// TIA Portal V17 export
// export: Created 2025-07-01T12:14:22.0161746Z, ExportSetting WithDefaults, DisplayName Totally Integrated Automation Portal, DisplayVersion V17, DisplayName TIA Portal Openness, DisplayVersion V17, DisplayName TIA Portal Version Control Interface, DisplayVersion V17, DisplayName SINAMICS Startdrive Advanced, DisplayVersion V17, DisplayName SINAMICS Startdrive G130, G150, S120, S150, SINAMICS MV, S210, DisplayVersion V17, DisplayName SINAMICS Startdrive G110M, G120, G120C, G120D, G120P, G115D, DisplayVersion V17, DisplayName STEP 7 Professional, DisplayVersion V17, DisplayName STEP 7 Safety, DisplayVersion V17, DisplayName WinCC Professional, DisplayVersion V17
FUNCTION_BLOCK "3PosLifter__Updated_V2_a4fa82_3a45ac7d-3c57-493c-83a9-58625a874be0 (2) - Copy_22ffb1"   // FB3, LAD
VERSION : 0.1
// stored: AutoNumber true, IsIECCheckEnabled false, UDAEnableTagReadback false
   VAR_INPUT
      iAreaClearConv : Bool;
      iAreaClearTransL2 : Bool;
      iAreaClear_TT : Bool;
      iAutoRunning : Bool;
      iErrorAck : Bool;
      iL1PalletPrsnt : Bool;
      iL1S1Raise : Bool;
      iL1S2Down : Bool;
      iL1S2DownOver : Bool;
      iL2PalletPrsent : Bool;
      iL2S1Down : Bool;
      iL2S1Raise : Bool;
      iL2s2DownOver : Bool;
      iL2s2Raise : Bool;
      iLiffterAtPos1 : Bool;
      iLiffterAtPos2 : Bool;
      iLiffterAtPos3 : Bool;
      iLiffterAtPos4 : Bool;
      iLifterAt1 : Bool;
      iLifterAtPos1 : Bool;
      iLifterAtPos2 : Bool;
      iLifterAtPos3 : Bool;
      iLifterAtPos4 : Bool;
      iOTSFrmConv : Bool;
      iPalAtTT : Bool;
      iPalletAtL1 : Bool;
      iPalletAtL2 : Bool;
      iPalletAtTT : Bool;
      iPalletPrsntL1 : Bool;
      iRTRFrmConv : Bool;
      iRTRFrmTT : Bool;
      iRTRFrm_TT : Bool;
      iReacvAreaClr : Bool;
      iReceiveAreaClear : Bool;
      iReceiveAreaClrConv : Bool;
      iRecvAreaClear : Bool;
      iReset_fault : Bool;
      iRunOutActive : Bool;
      iRunOutCycle : Bool;
      iSstMode : Bool;
      iSstPB : Bool;
      iTransAreaClearConv : Bool;
      iTransAreaClr : Bool;
      ipalletPrsntAtTT : Bool;
   END_VAR
   VAR_OUTPUT
      qL1S1Down : Bool;
      qL1S1raise : Bool;
      qL1S2Down : Bool;
      qL1S2Raise : Bool;
      qL1TrnsfrConv : Bool;
      qL2S1raise : Bool;
      qL2S2Down : Bool;
      qL2S2Raise : Bool;
      qLiffterAtPos2 : Bool;
      qLifterAtPos1 : Bool;
      qLifterAtPos3 : Bool;
      qLifterAtPos4 : Bool;
      qLifterGotoPos1 : Bool;
      qOTSToNext : Bool;
      qOTSTo_TT : Bool;
      qOutput1 : Bool;
      qRTRToConv : Bool;
      qRTRToTT : Bool;
      qRTR_To_Conv : Bool;
   END_VAR
   VAR_IN_OUT
      IqRx_Frm_TT : Bool;
      iqRx_frm_Conv : Bool;
      iqTX_To_Conv : Bool;
      iqTX_To_TT : Bool;
      iqTx_To_ConvPos4 : Bool;
      iqTx_To_Rej : Bool;
   END_VAR
   VAR DB_SPECIFIC
      StateNo : Int;
      s190_sStWtL1RcvComplete_T1 : Bool;
      s200_sStWtForL1StprUp_T1 : Bool;
      s240_sStWtL2TransComplete_T1 : Bool;
      s250_sStWtDeforkDone : Bool;
      s250_sStWtDeforkDone_Cond1 : Bool;
      s250_sStWtDeforkDone_Cond2 : Bool;
      s250_sStWtDeforkDone_T1 : Bool;
      sInitialConvRun : Bool;
      sInitialConvRun_T1 : Bool;
      sOTSTimeout : Bool;
      sSeq1Over : Bool;
      sSeq2Over : Bool;
      sSst : Bool;
      sSstPulse : Bool;
      sSstRise : Bool;
      sStChkPalAtTT : Bool;
      sStChkPalAtTT_T1 : Bool;
      sStChkPalAtTT_T2 : Bool;
      sStChkPalAtTT_T3 : Bool;
      sStChkPalletAtTT : Bool;
      sStChkPalletAtTT1 : Bool;
      sStChkPalletAtTT1_T1 : Bool;
      sStChkPalletAtTT1_T2 : Bool;
      sStChkPalletAtTT_T1 : Bool;
      sStChkPalletAtTT_T2 : Bool;
      sStChkPalletPrsntL1L2 : Bool;
      sStChkPalletPrsntL1L2_T1 : Bool;
      sStChkPalletPrsntL1L2_T2 : Bool;
      sStChkPalletPrsntL1L2_T3 : Bool;
      sStChkPalletPrsntL1L2_T4 : Bool;
      sStChkRunOutActive1 : Bool;
      sStChkRunOutActive1_T1 : Bool;
      sStChkRunOutActive1_T2 : Bool;
      sStL1S2Down : Bool;
      sStL1S2DownOver : Bool;
      sStL1S2DownOver_T1 : Bool;
      sStL1S2Down_T1 : Bool;
      sStNextRdyInTransit : Bool;
      sStNextRdyInTransit_1 : Bool;
      sStNextRdyInTransit_1_T1 : Bool;
      sStNextRdyInTransit_1_T2 : Bool;
      sStNextRdyInTransit_3 : Bool;
      sStNextRdyInTransit_3_T1 : Bool;
      sStNextRdyInTransit_3_T2 : Bool;
      sStNextRdyInTransit_T1 : Bool;
      sStNextRdyInTransit_T2 : Bool;
      sStRecovery : Bool;
      sStRecovery_T1 : Bool;
      sStRecovery_T2 : Bool;
      sStRecovery_T3 : Bool;
      sStRecovery_T4 : Bool;
      sStRecovery_T5 : Bool;
      sStRecovery_T6 : Bool;
      sStRecovery_T7 : Bool;
      sStRecovery_T8 : Bool;
      sStRunOutActive : Bool;
      sStRunOutActive_T1 : Bool;
      sStRunOutActive_T2 : Bool;
      sStWtDeforkDone : Bool;
      sStWtDeforkDone_T1 : Bool;
      sStWtForFaultReset : Bool;
      sStWtForFaultReset_T1 : Bool;
      sStWtForL1L2StoprsUp : Bool;
      sStWtForL1L2StoprsUp_T1 : Bool;
      sStWtForL1StprUp : Bool;
      sStWtForL1StprUp_T1 : Bool;
      sStWtL1PalRcvDone : Bool;
      sStWtL1PalRcvDone_T1 : Bool;
      sStWtL1RcvComplete : Bool;
      sStWtL1RcvComplete_T1 : Bool;
      sStWtL1RecvBegin : Bool;
      sStWtL1RecvBegin_T1 : Bool;
      sStWtL1S1Down1 : Bool;
      sStWtL1S1Down1_T1 : Bool;
      sStWtL1S2DownOver : Bool;
      sStWtL1S2DownOver_T1 : Bool;
      sStWtL1TransBegin : Bool;
      sStWtL1TransBeginPos4 : Bool;
      sStWtL1TransBeginPos4_T1 : Bool;
      sStWtL1TransBegin_T1 : Bool;
      sStWtL1TransComplet : Bool;
      sStWtL1TransComplet_T1 : Bool;
      sStWtL2RcvDone : Bool;
      sStWtL2RcvDone_T1 : Bool;
      sStWtL2RecvingActive : Bool;
      sStWtL2RecvingActive_T1 : Bool;
      sStWtL2S1Down : Bool;
      sStWtL2S1Down_T1 : Bool;
      sStWtL2S2Down : Bool;
      sStWtL2S2Down_T1 : Bool;
      sStWtL2TranBegin : Bool;
      sStWtL2TranBegin_T1 : Bool;
      sStWtL2TransComplete : Bool;
      sStWtL2TransComplete_T1 : Bool;
      sStWtLifterAtPos1 : Bool;
      sStWtLifterAtPos1_T1 : Bool;
      sStWtLifterAtPos2 : Bool;
      sStWtLifterAtPos2_T1 : Bool;
      sStWtLifterAtPos3 : Bool;
      sStWtLifterAtPos3_T1 : Bool;
      sStWtLifterAtPos4 : Bool;
      sStWtLifterAtPos4_T1 : Bool;
      sStWtLifterAtPosn1 : Bool;
      sStWtLifterAtPosn1_T1 : Bool;
      sStWtOTSFrmConv : Bool;
      sStWtOTSFrmConv1 : Bool;
      sStWtOTSFrmConv1_T1 : Bool;
      sStWtOTSFrmConv1_T2 : Bool;
      sStWtOTSFrmConv_T1 : Bool;
      sStWtOTSFrmTT : Bool;
      sStWtOTSFrmTT_T1 : Bool;
      sStWtRTRFrmConvPos4 : Bool;
      sStWtRTRFrmConvPos4_T1 : Bool;
      sStWtRTRFrmTT : Bool;
      sStWtRTRFrmTT_T1 : Bool;
      sStWtRcvBegin : Bool;
      sStWtRcvBegin_T1 : Bool;
      sStWtResetRel : Bool;
      sStWtResetRel_T1 : Bool;
      sStWtTransDonePos4 : Bool;
      sStWtTransDonePos4_T1 : Bool;
   END_VAR
   VAR_TEMP
      tOne : Bool;
   END_VAR
   VAR_TEMP   // added for the SCL form of the ladder/FBD networks
      _w1 : Bool;
   END_VAR
BEGIN

REGION Network 1
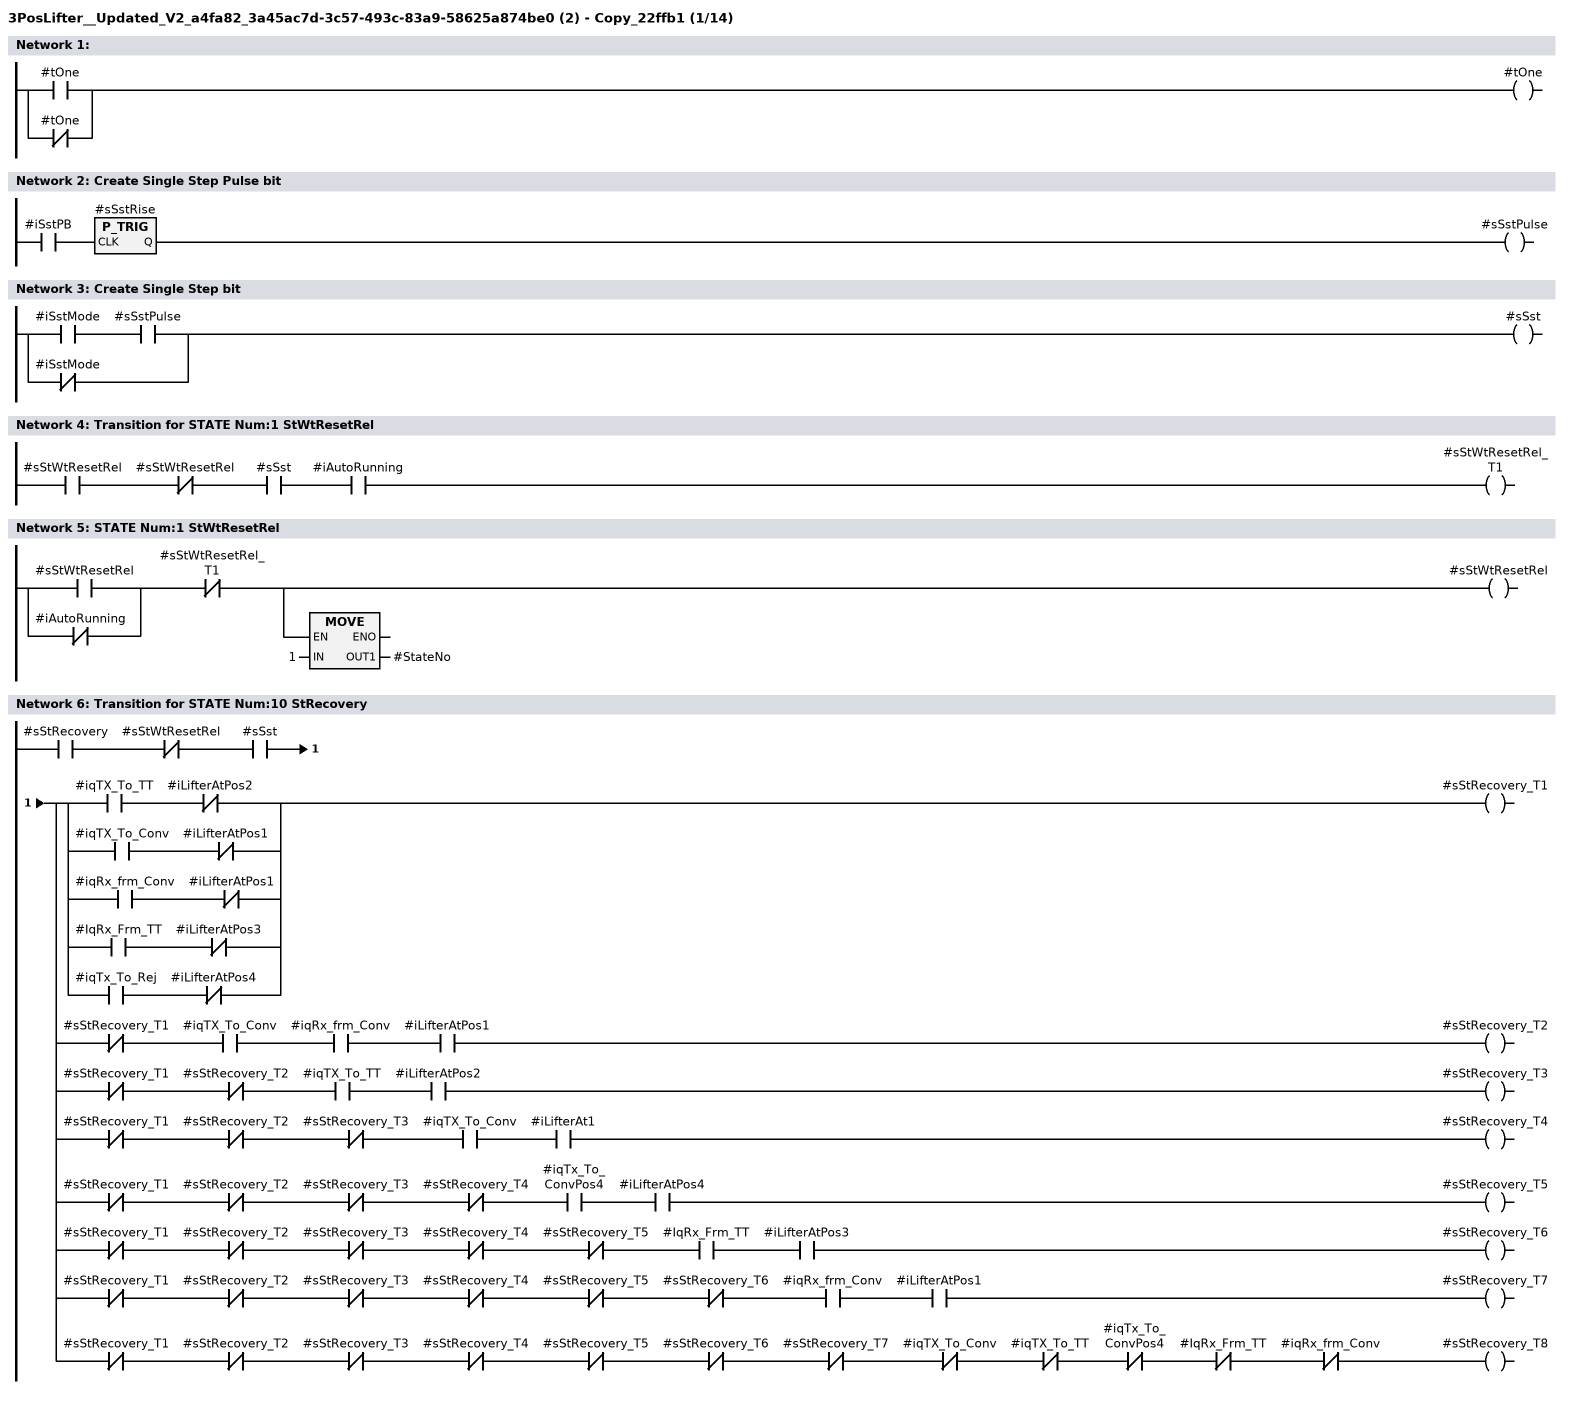
   RUNG wire#powerrail
      Contact( #tOne )
      wire#w1
      Coil( #tOne )
   END_RUNG
   RUNG wire#powerrail
      I_Contact( #tOne )
   END_RUNG wire#w1
   // the same network as SCL:
   #tOne := #tOne OR NOT #tOne;
END_REGION

REGION Network 2: Create Single Step Pulse bit
   RUNG wire#powerrail
      Contact( #iSstPB )
      P_Trig( #sSstRise )
      Coil( #sSstPulse )
   END_RUNG
   // the same network as SCL:
   #_w1 := #iSstPB AND NOT #sSstRise;   // rising edge
   #sSstRise := #iSstPB;
   #sSstPulse := #_w1;
END_REGION

REGION Network 3: Create Single Step bit
   RUNG wire#powerrail
      Contact( #iSstMode )
      Contact( #sSstPulse )
      wire#w1
      Coil( #sSst )
   END_RUNG
   RUNG wire#powerrail
      I_Contact( #iSstMode )
   END_RUNG wire#w1
   // the same network as SCL:
   #sSst := (#iSstMode AND #sSstPulse) OR NOT #iSstMode;
END_REGION

REGION Network 4: Transition for STATE Num:1 StWtResetRel
   RUNG wire#powerrail
      Contact( #sStWtResetRel )
      I_Contact( #sStWtResetRel )
      Contact( #sSst )
      Contact( #iAutoRunning )
      Coil( #sStWtResetRel_T1 )
   END_RUNG
   // the same network as SCL:
   #sStWtResetRel_T1 := #sStWtResetRel AND NOT #sStWtResetRel AND #sSst AND #iAutoRunning;
END_REGION

REGION Network 5: STATE Num:1 StWtResetRel
   RUNG wire#powerrail
      Contact( #sStWtResetRel )
      wire#w1
      I_Contact( #sStWtResetRel_T1 )
      wire#w2
      Coil( #sStWtResetRel )
   END_RUNG
   RUNG wire#powerrail
      I_Contact( #iAutoRunning )
   END_RUNG wire#w1
   RUNG wire#w2
      { S7_GenerateENO := "TRUE" } Move(in := 1, out1 => #StateNo)
   END_RUNG
   // the same network as SCL:
   #sStWtResetRel := (#sStWtResetRel OR NOT #iAutoRunning) AND NOT #sStWtResetRel_T1;
   IF #sStWtResetRel THEN #StateNo := 1; END_IF;
END_REGION

REGION Network 6: Transition for STATE Num:10 StRecovery
   RUNG wire#powerrail
      Contact( #sStRecovery )
      I_Contact( #sStWtResetRel )
      Contact( #sSst )
      wire#w1
      Contact( #iqTX_To_TT )
      I_Contact( #iLifterAtPos2 )
      wire#w2
      Coil( #sStRecovery_T1 )
   END_RUNG
   RUNG wire#w1
      Contact( #iqTX_To_Conv )
      I_Contact( #iLifterAtPos1 )
   END_RUNG wire#w2
   RUNG wire#w1
      Contact( #iqRx_frm_Conv )
      I_Contact( #iLifterAtPos1 )
   END_RUNG wire#w2
   RUNG wire#w1
      Contact( #IqRx_Frm_TT )
      I_Contact( #iLifterAtPos3 )
   END_RUNG wire#w2
   RUNG wire#w1
      Contact( #iqTx_To_Rej )
      I_Contact( #iLifterAtPos4 )
   END_RUNG wire#w2
   RUNG wire#w1
      I_Contact( #sStRecovery_T1 )
      Contact( #iqTX_To_Conv )
      Contact( #iqRx_frm_Conv )
      Contact( #iLifterAtPos1 )
      Coil( #sStRecovery_T2 )
   END_RUNG
   RUNG wire#w1
      I_Contact( #sStRecovery_T1 )
      I_Contact( #sStRecovery_T2 )
      Contact( #iqTX_To_TT )
      Contact( #iLifterAtPos2 )
      Coil( #sStRecovery_T3 )
   END_RUNG
   RUNG wire#w1
      I_Contact( #sStRecovery_T1 )
      I_Contact( #sStRecovery_T2 )
      I_Contact( #sStRecovery_T3 )
      Contact( #iqTX_To_Conv )
      Contact( #iLifterAt1 )
      Coil( #sStRecovery_T4 )
   END_RUNG
   RUNG wire#w1
      I_Contact( #sStRecovery_T1 )
      I_Contact( #sStRecovery_T2 )
      I_Contact( #sStRecovery_T3 )
      I_Contact( #sStRecovery_T4 )
      Contact( #iqTx_To_ConvPos4 )
      Contact( #iLifterAtPos4 )
      Coil( #sStRecovery_T5 )
   END_RUNG
   RUNG wire#w1
      I_Contact( #sStRecovery_T1 )
      I_Contact( #sStRecovery_T2 )
      I_Contact( #sStRecovery_T3 )
      I_Contact( #sStRecovery_T4 )
      I_Contact( #sStRecovery_T5 )
      Contact( #IqRx_Frm_TT )
      Contact( #iLifterAtPos3 )
      Coil( #sStRecovery_T6 )
   END_RUNG
   RUNG wire#w1
      I_Contact( #sStRecovery_T1 )
      I_Contact( #sStRecovery_T2 )
      I_Contact( #sStRecovery_T3 )
      I_Contact( #sStRecovery_T4 )
      I_Contact( #sStRecovery_T5 )
      I_Contact( #sStRecovery_T6 )
      Contact( #iqRx_frm_Conv )
      Contact( #iLifterAtPos1 )
      Coil( #sStRecovery_T7 )
   END_RUNG
   RUNG wire#w1
      I_Contact( #sStRecovery_T1 )
      I_Contact( #sStRecovery_T2 )
      I_Contact( #sStRecovery_T3 )
      I_Contact( #sStRecovery_T4 )
      I_Contact( #sStRecovery_T5 )
      I_Contact( #sStRecovery_T6 )
      I_Contact( #sStRecovery_T7 )
      I_Contact( #iqTX_To_Conv )
      I_Contact( #iqTX_To_TT )
      I_Contact( #iqTx_To_ConvPos4 )
      I_Contact( #IqRx_Frm_TT )
      I_Contact( #iqRx_frm_Conv )
      Coil( #sStRecovery_T8 )
   END_RUNG
   // the same network as SCL:
   #_w1 := #sStRecovery AND NOT #sStWtResetRel AND #sSst;
   #sStRecovery_T1 := #_w1 AND ((#iqTX_To_TT AND NOT #iLifterAtPos2) OR (#iqTX_To_Conv AND NOT #iLifterAtPos1) OR (#iqRx_frm_Conv AND NOT #iLifterAtPos1) OR (#IqRx_Frm_TT AND NOT #iLifterAtPos3) OR (#iqTx_To_Rej AND NOT #iLifterAtPos4));
   #sStRecovery_T2 := #_w1 AND NOT #sStRecovery_T1 AND #iqTX_To_Conv AND #iqRx_frm_Conv AND #iLifterAtPos1;
   #sStRecovery_T3 := #_w1 AND NOT #sStRecovery_T1 AND NOT #sStRecovery_T2 AND #iqTX_To_TT AND #iLifterAtPos2;
   #sStRecovery_T4 := #_w1 AND NOT #sStRecovery_T1 AND NOT #sStRecovery_T2 AND NOT #sStRecovery_T3 AND #iqTX_To_Conv AND #iLifterAt1;
   #sStRecovery_T5 := #_w1 AND NOT #sStRecovery_T1 AND NOT #sStRecovery_T2 AND NOT #sStRecovery_T3 AND NOT #sStRecovery_T4 AND #iqTx_To_ConvPos4 AND #iLifterAtPos4;
   #sStRecovery_T6 := #_w1 AND NOT #sStRecovery_T1 AND NOT #sStRecovery_T2 AND NOT #sStRecovery_T3 AND NOT #sStRecovery_T4 AND NOT #sStRecovery_T5 AND #IqRx_Frm_TT AND #iLifterAtPos3;
   #sStRecovery_T7 := #_w1 AND NOT #sStRecovery_T1 AND NOT #sStRecovery_T2 AND NOT #sStRecovery_T3 AND NOT #sStRecovery_T4 AND NOT #sStRecovery_T5 AND NOT #sStRecovery_T6 AND #iqRx_frm_Conv AND #iLifterAtPos1;
   #sStRecovery_T8 := #_w1 AND NOT #sStRecovery_T1 AND NOT #sStRecovery_T2 AND NOT #sStRecovery_T3 AND NOT #sStRecovery_T4 AND NOT #sStRecovery_T5 AND NOT #sStRecovery_T6 AND NOT #sStRecovery_T7 AND NOT #iqTX_To_Conv AND NOT #iqTX_To_TT AND NOT #iqTx_To_ConvPos4 AND NOT #IqRx_Frm_TT AND NOT #iqRx_frm_Conv;
END_REGION

REGION Network 7: STATE Num:10 StRecovery
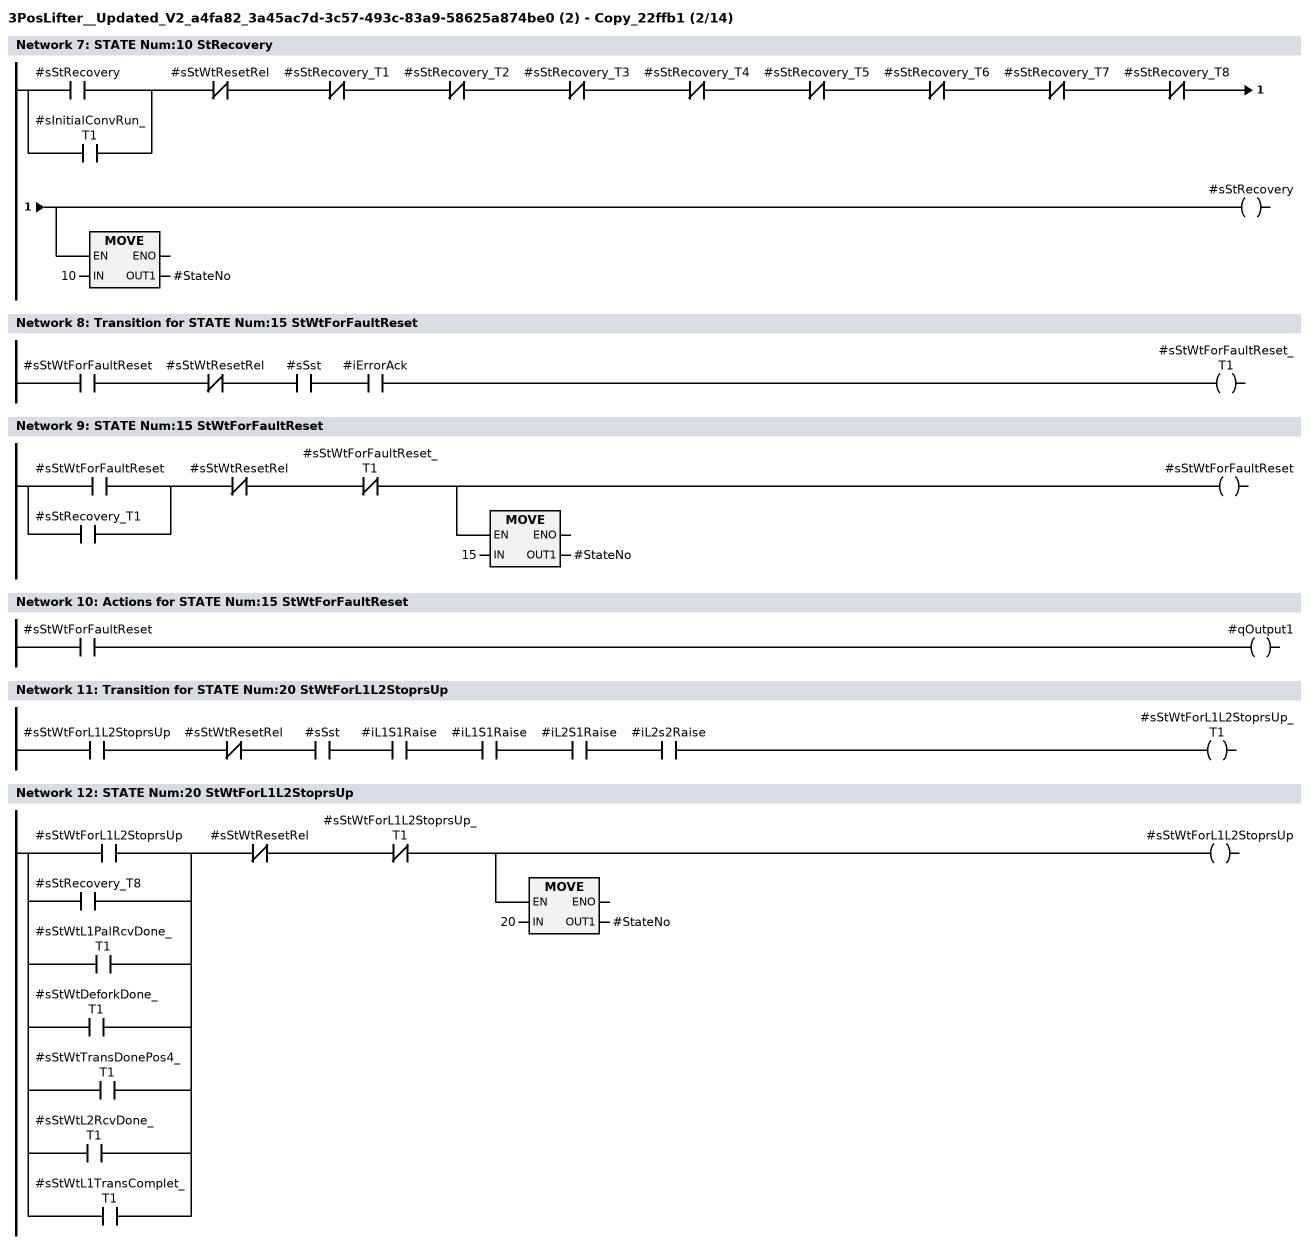
   RUNG wire#powerrail
      Contact( #sStRecovery )
      wire#w1
      I_Contact( #sStWtResetRel )
      I_Contact( #sStRecovery_T1 )
      I_Contact( #sStRecovery_T2 )
      I_Contact( #sStRecovery_T3 )
      I_Contact( #sStRecovery_T4 )
      I_Contact( #sStRecovery_T5 )
      I_Contact( #sStRecovery_T6 )
      I_Contact( #sStRecovery_T7 )
      I_Contact( #sStRecovery_T8 )
      wire#w2
      Coil( #sStRecovery )
   END_RUNG
   RUNG wire#powerrail
      Contact( #sInitialConvRun_T1 )
   END_RUNG wire#w1
   RUNG wire#w2
      { S7_GenerateENO := "TRUE" } Move(in := 10, out1 => #StateNo)
   END_RUNG
   // the same network as SCL:
   #sStRecovery := (#sStRecovery OR #sInitialConvRun_T1) AND NOT #sStWtResetRel AND NOT #sStRecovery_T1 AND NOT #sStRecovery_T2 AND NOT #sStRecovery_T3 AND NOT #sStRecovery_T4 AND NOT #sStRecovery_T5 AND NOT #sStRecovery_T6 AND NOT #sStRecovery_T7 AND NOT #sStRecovery_T8;
   IF #sStRecovery THEN #StateNo := 10; END_IF;
END_REGION

REGION Network 8: Transition for STATE Num:15 StWtForFaultReset
   RUNG wire#powerrail
      Contact( #sStWtForFaultReset )
      I_Contact( #sStWtResetRel )
      Contact( #sSst )
      Contact( #iErrorAck )
      Coil( #sStWtForFaultReset_T1 )
   END_RUNG
   // the same network as SCL:
   #sStWtForFaultReset_T1 := #sStWtForFaultReset AND NOT #sStWtResetRel AND #sSst AND #iErrorAck;
END_REGION

REGION Network 9: STATE Num:15 StWtForFaultReset
   RUNG wire#powerrail
      Contact( #sStWtForFaultReset )
      wire#w1
      I_Contact( #sStWtResetRel )
      I_Contact( #sStWtForFaultReset_T1 )
      wire#w2
      Coil( #sStWtForFaultReset )
   END_RUNG
   RUNG wire#powerrail
      Contact( #sStRecovery_T1 )
   END_RUNG wire#w1
   RUNG wire#w2
      { S7_GenerateENO := "TRUE" } Move(in := 15, out1 => #StateNo)
   END_RUNG
   // the same network as SCL:
   #sStWtForFaultReset := (#sStWtForFaultReset OR #sStRecovery_T1) AND NOT #sStWtResetRel AND NOT #sStWtForFaultReset_T1;
   IF #sStWtForFaultReset THEN #StateNo := 15; END_IF;
END_REGION

REGION Network 10: Actions for STATE Num:15 StWtForFaultReset
   RUNG wire#powerrail
      Contact( #sStWtForFaultReset )
      Coil( #qOutput1 )
   END_RUNG
   // the same network as SCL:
   #qOutput1 := #sStWtForFaultReset;
END_REGION

REGION Network 11: Transition for STATE Num:20 StWtForL1L2StoprsUp
   RUNG wire#powerrail
      Contact( #sStWtForL1L2StoprsUp )
      I_Contact( #sStWtResetRel )
      Contact( #sSst )
      Contact( #iL1S1Raise )
      Contact( #iL1S1Raise )
      Contact( #iL2S1Raise )
      Contact( #iL2s2Raise )
      Coil( #sStWtForL1L2StoprsUp_T1 )
   END_RUNG
   // the same network as SCL:
   #sStWtForL1L2StoprsUp_T1 := #sStWtForL1L2StoprsUp AND NOT #sStWtResetRel AND #sSst AND #iL1S1Raise AND #iL1S1Raise AND #iL2S1Raise AND #iL2s2Raise;
END_REGION

REGION Network 12: STATE Num:20 StWtForL1L2StoprsUp
   RUNG wire#powerrail
      Contact( #sStWtForL1L2StoprsUp )
      wire#w1
      I_Contact( #sStWtResetRel )
      I_Contact( #sStWtForL1L2StoprsUp_T1 )
      wire#w2
      Coil( #sStWtForL1L2StoprsUp )
   END_RUNG
   RUNG wire#powerrail
      Contact( #sStRecovery_T8 )
   END_RUNG wire#w1
   RUNG wire#powerrail
      Contact( #sStWtL1PalRcvDone_T1 )
   END_RUNG wire#w1
   RUNG wire#powerrail
      Contact( #sStWtDeforkDone_T1 )
   END_RUNG wire#w1
   RUNG wire#powerrail
      Contact( #sStWtTransDonePos4_T1 )
   END_RUNG wire#w1
   RUNG wire#powerrail
      Contact( #sStWtL2RcvDone_T1 )
   END_RUNG wire#w1
   RUNG wire#powerrail
      Contact( #sStWtL1TransComplet_T1 )
   END_RUNG wire#w1
   RUNG wire#w2
      { S7_GenerateENO := "TRUE" } Move(in := 20, out1 => #StateNo)
   END_RUNG
   // the same network as SCL:
   #sStWtForL1L2StoprsUp := (#sStWtForL1L2StoprsUp OR #sStRecovery_T8 OR #sStWtL1PalRcvDone_T1 OR #sStWtDeforkDone_T1 OR #sStWtTransDonePos4_T1 OR #sStWtL2RcvDone_T1 OR #sStWtL1TransComplet_T1) AND NOT #sStWtResetRel AND NOT #sStWtForL1L2StoprsUp_T1;
   IF #sStWtForL1L2StoprsUp THEN #StateNo := 20; END_IF;
END_REGION

REGION Network 13: Actions for STATE Num:20 StWtForL1L2StoprsUp
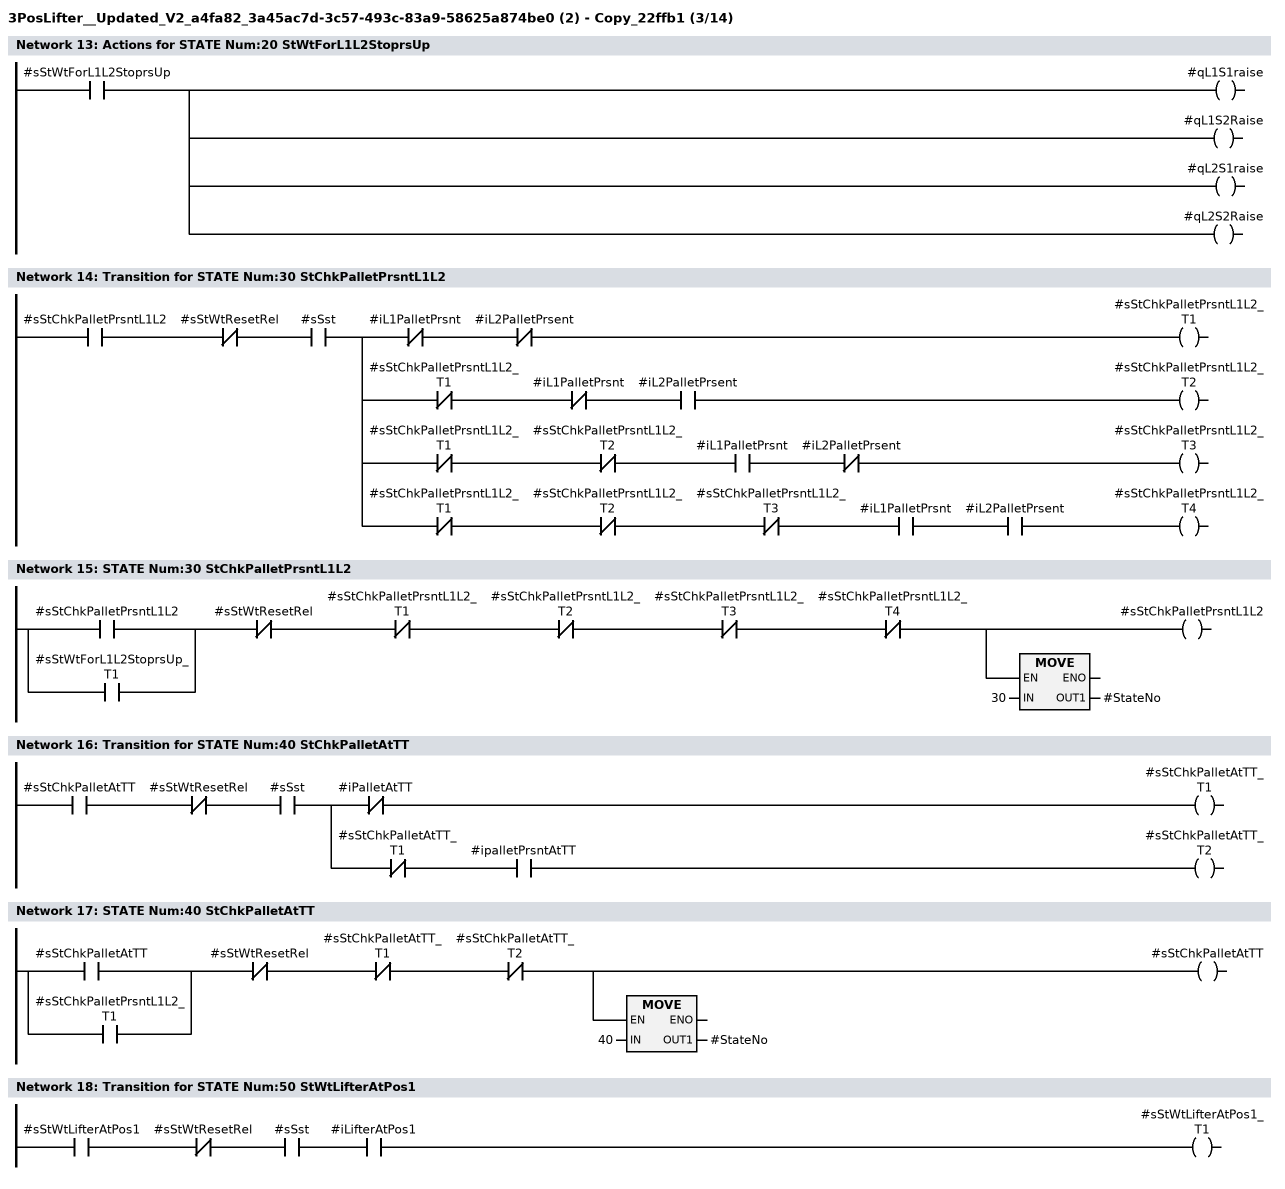
   RUNG wire#powerrail
      Contact( #sStWtForL1L2StoprsUp )
      wire#w1
      Coil( #qL1S1raise )
   END_RUNG
   RUNG wire#w1
      Coil( #qL1S2Raise )
   END_RUNG
   RUNG wire#w1
      Coil( #qL2S1raise )
   END_RUNG
   RUNG wire#w1
      Coil( #qL2S2Raise )
   END_RUNG
   // the same network as SCL:
   #qL1S1raise := #sStWtForL1L2StoprsUp;
   #qL1S2Raise := #sStWtForL1L2StoprsUp;
   #qL2S1raise := #sStWtForL1L2StoprsUp;
   #qL2S2Raise := #sStWtForL1L2StoprsUp;
END_REGION

REGION Network 14: Transition for STATE Num:30 StChkPalletPrsntL1L2
   RUNG wire#powerrail
      Contact( #sStChkPalletPrsntL1L2 )
      I_Contact( #sStWtResetRel )
      Contact( #sSst )
      wire#w1
      I_Contact( #iL1PalletPrsnt )
      I_Contact( #iL2PalletPrsent )
      Coil( #sStChkPalletPrsntL1L2_T1 )
   END_RUNG
   RUNG wire#w1
      I_Contact( #sStChkPalletPrsntL1L2_T1 )
      I_Contact( #iL1PalletPrsnt )
      Contact( #iL2PalletPrsent )
      Coil( #sStChkPalletPrsntL1L2_T2 )
   END_RUNG
   RUNG wire#w1
      I_Contact( #sStChkPalletPrsntL1L2_T1 )
      I_Contact( #sStChkPalletPrsntL1L2_T2 )
      Contact( #iL1PalletPrsnt )
      I_Contact( #iL2PalletPrsent )
      Coil( #sStChkPalletPrsntL1L2_T3 )
   END_RUNG
   RUNG wire#w1
      I_Contact( #sStChkPalletPrsntL1L2_T1 )
      I_Contact( #sStChkPalletPrsntL1L2_T2 )
      I_Contact( #sStChkPalletPrsntL1L2_T3 )
      Contact( #iL1PalletPrsnt )
      Contact( #iL2PalletPrsent )
      Coil( #sStChkPalletPrsntL1L2_T4 )
   END_RUNG
   // the same network as SCL:
   #_w1 := #sStChkPalletPrsntL1L2 AND NOT #sStWtResetRel AND #sSst;
   #sStChkPalletPrsntL1L2_T1 := #_w1 AND NOT #iL1PalletPrsnt AND NOT #iL2PalletPrsent;
   #sStChkPalletPrsntL1L2_T2 := #_w1 AND NOT #sStChkPalletPrsntL1L2_T1 AND NOT #iL1PalletPrsnt AND #iL2PalletPrsent;
   #sStChkPalletPrsntL1L2_T3 := #_w1 AND NOT #sStChkPalletPrsntL1L2_T1 AND NOT #sStChkPalletPrsntL1L2_T2 AND #iL1PalletPrsnt AND NOT #iL2PalletPrsent;
   #sStChkPalletPrsntL1L2_T4 := #_w1 AND NOT #sStChkPalletPrsntL1L2_T1 AND NOT #sStChkPalletPrsntL1L2_T2 AND NOT #sStChkPalletPrsntL1L2_T3 AND #iL1PalletPrsnt AND #iL2PalletPrsent;
END_REGION

REGION Network 15: STATE Num:30 StChkPalletPrsntL1L2
   RUNG wire#powerrail
      Contact( #sStChkPalletPrsntL1L2 )
      wire#w1
      I_Contact( #sStWtResetRel )
      I_Contact( #sStChkPalletPrsntL1L2_T1 )
      I_Contact( #sStChkPalletPrsntL1L2_T2 )
      I_Contact( #sStChkPalletPrsntL1L2_T3 )
      I_Contact( #sStChkPalletPrsntL1L2_T4 )
      wire#w2
      Coil( #sStChkPalletPrsntL1L2 )
   END_RUNG
   RUNG wire#powerrail
      Contact( #sStWtForL1L2StoprsUp_T1 )
   END_RUNG wire#w1
   RUNG wire#w2
      { S7_GenerateENO := "TRUE" } Move(in := 30, out1 => #StateNo)
   END_RUNG
   // the same network as SCL:
   #sStChkPalletPrsntL1L2 := (#sStChkPalletPrsntL1L2 OR #sStWtForL1L2StoprsUp_T1) AND NOT #sStWtResetRel AND NOT #sStChkPalletPrsntL1L2_T1 AND NOT #sStChkPalletPrsntL1L2_T2 AND NOT #sStChkPalletPrsntL1L2_T3 AND NOT #sStChkPalletPrsntL1L2_T4;
   IF #sStChkPalletPrsntL1L2 THEN #StateNo := 30; END_IF;
END_REGION

REGION Network 16: Transition for STATE Num:40 StChkPalletAtTT
   RUNG wire#powerrail
      Contact( #sStChkPalletAtTT )
      I_Contact( #sStWtResetRel )
      Contact( #sSst )
      wire#w1
      I_Contact( #iPalletAtTT )
      Coil( #sStChkPalletAtTT_T1 )
   END_RUNG
   RUNG wire#w1
      I_Contact( #sStChkPalletAtTT_T1 )
      Contact( #ipalletPrsntAtTT )
      Coil( #sStChkPalletAtTT_T2 )
   END_RUNG
   // the same network as SCL:
   #_w1 := #sStChkPalletAtTT AND NOT #sStWtResetRel AND #sSst;
   #sStChkPalletAtTT_T1 := #_w1 AND NOT #iPalletAtTT;
   #sStChkPalletAtTT_T2 := #_w1 AND NOT #sStChkPalletAtTT_T1 AND #ipalletPrsntAtTT;
END_REGION

REGION Network 17: STATE Num:40 StChkPalletAtTT
   RUNG wire#powerrail
      Contact( #sStChkPalletAtTT )
      wire#w1
      I_Contact( #sStWtResetRel )
      I_Contact( #sStChkPalletAtTT_T1 )
      I_Contact( #sStChkPalletAtTT_T2 )
      wire#w2
      Coil( #sStChkPalletAtTT )
   END_RUNG
   RUNG wire#powerrail
      Contact( #sStChkPalletPrsntL1L2_T1 )
   END_RUNG wire#w1
   RUNG wire#w2
      { S7_GenerateENO := "TRUE" } Move(in := 40, out1 => #StateNo)
   END_RUNG
   // the same network as SCL:
   #sStChkPalletAtTT := (#sStChkPalletAtTT OR #sStChkPalletPrsntL1L2_T1) AND NOT #sStWtResetRel AND NOT #sStChkPalletAtTT_T1 AND NOT #sStChkPalletAtTT_T2;
   IF #sStChkPalletAtTT THEN #StateNo := 40; END_IF;
END_REGION

REGION Network 18: Transition for STATE Num:50 StWtLifterAtPos1
   RUNG wire#powerrail
      Contact( #sStWtLifterAtPos1 )
      I_Contact( #sStWtResetRel )
      Contact( #sSst )
      Contact( #iLifterAtPos1 )
      Coil( #sStWtLifterAtPos1_T1 )
   END_RUNG
   // the same network as SCL:
   #sStWtLifterAtPos1_T1 := #sStWtLifterAtPos1 AND NOT #sStWtResetRel AND #sSst AND #iLifterAtPos1;
END_REGION

REGION Network 19: STATE Num:50 StWtLifterAtPos1
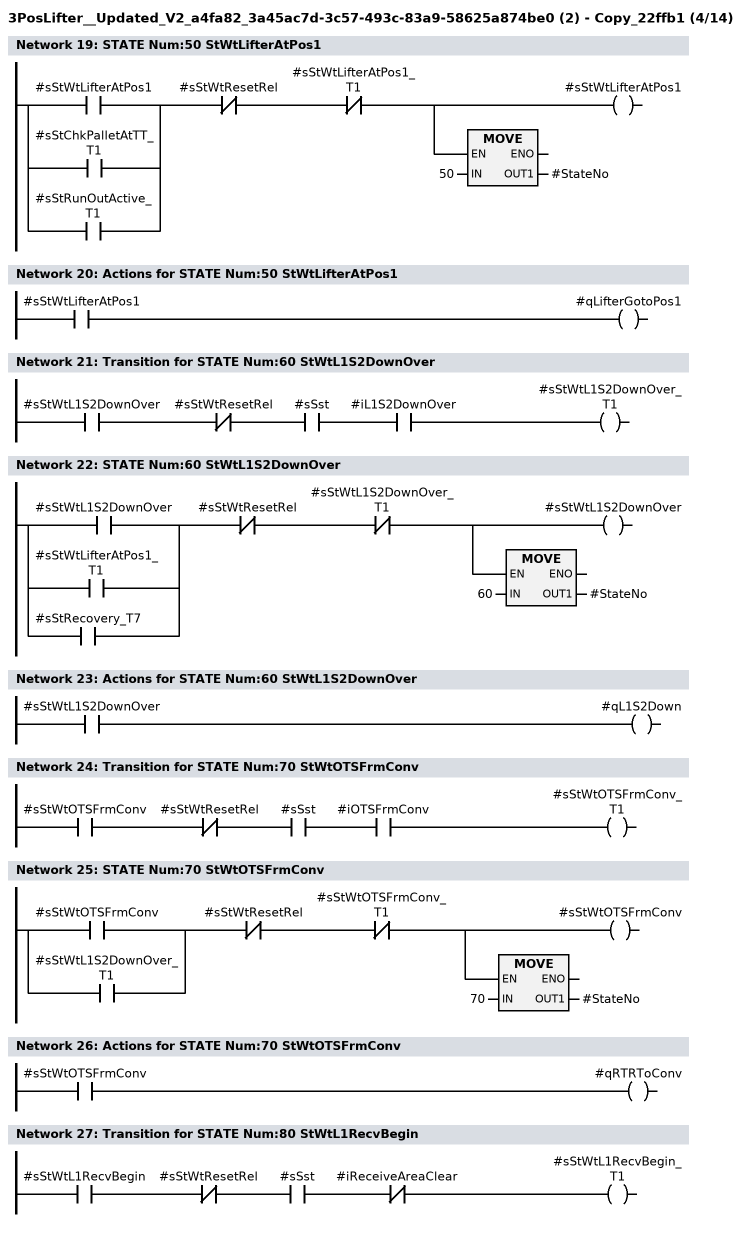
   RUNG wire#powerrail
      Contact( #sStWtLifterAtPos1 )
      wire#w1
      I_Contact( #sStWtResetRel )
      I_Contact( #sStWtLifterAtPos1_T1 )
      wire#w2
      Coil( #sStWtLifterAtPos1 )
   END_RUNG
   RUNG wire#powerrail
      Contact( #sStChkPalletAtTT_T1 )
   END_RUNG wire#w1
   RUNG wire#powerrail
      Contact( #sStRunOutActive_T1 )
   END_RUNG wire#w1
   RUNG wire#w2
      { S7_GenerateENO := "TRUE" } Move(in := 50, out1 => #StateNo)
   END_RUNG
   // the same network as SCL:
   #sStWtLifterAtPos1 := (#sStWtLifterAtPos1 OR #sStChkPalletAtTT_T1 OR #sStRunOutActive_T1) AND NOT #sStWtResetRel AND NOT #sStWtLifterAtPos1_T1;
   IF #sStWtLifterAtPos1 THEN #StateNo := 50; END_IF;
END_REGION

REGION Network 20: Actions for STATE Num:50 StWtLifterAtPos1
   RUNG wire#powerrail
      Contact( #sStWtLifterAtPos1 )
      Coil( #qLifterGotoPos1 )
   END_RUNG
   // the same network as SCL:
   #qLifterGotoPos1 := #sStWtLifterAtPos1;
END_REGION

REGION Network 21: Transition for STATE Num:60 StWtL1S2DownOver
   RUNG wire#powerrail
      Contact( #sStWtL1S2DownOver )
      I_Contact( #sStWtResetRel )
      Contact( #sSst )
      Contact( #iL1S2DownOver )
      Coil( #sStWtL1S2DownOver_T1 )
   END_RUNG
   // the same network as SCL:
   #sStWtL1S2DownOver_T1 := #sStWtL1S2DownOver AND NOT #sStWtResetRel AND #sSst AND #iL1S2DownOver;
END_REGION

REGION Network 22: STATE Num:60 StWtL1S2DownOver
   RUNG wire#powerrail
      Contact( #sStWtL1S2DownOver )
      wire#w1
      I_Contact( #sStWtResetRel )
      I_Contact( #sStWtL1S2DownOver_T1 )
      wire#w2
      Coil( #sStWtL1S2DownOver )
   END_RUNG
   RUNG wire#powerrail
      Contact( #sStWtLifterAtPos1_T1 )
   END_RUNG wire#w1
   RUNG wire#powerrail
      Contact( #sStRecovery_T7 )
   END_RUNG wire#w1
   RUNG wire#w2
      { S7_GenerateENO := "TRUE" } Move(in := 60, out1 => #StateNo)
   END_RUNG
   // the same network as SCL:
   #sStWtL1S2DownOver := (#sStWtL1S2DownOver OR #sStWtLifterAtPos1_T1 OR #sStRecovery_T7) AND NOT #sStWtResetRel AND NOT #sStWtL1S2DownOver_T1;
   IF #sStWtL1S2DownOver THEN #StateNo := 60; END_IF;
END_REGION

REGION Network 23: Actions for STATE Num:60 StWtL1S2DownOver
   RUNG wire#powerrail
      Contact( #sStWtL1S2DownOver )
      Coil( #qL1S2Down )
   END_RUNG
   // the same network as SCL:
   #qL1S2Down := #sStWtL1S2DownOver;
END_REGION

REGION Network 24: Transition for STATE Num:70 StWtOTSFrmConv
   RUNG wire#powerrail
      Contact( #sStWtOTSFrmConv )
      I_Contact( #sStWtResetRel )
      Contact( #sSst )
      Contact( #iOTSFrmConv )
      Coil( #sStWtOTSFrmConv_T1 )
   END_RUNG
   // the same network as SCL:
   #sStWtOTSFrmConv_T1 := #sStWtOTSFrmConv AND NOT #sStWtResetRel AND #sSst AND #iOTSFrmConv;
END_REGION

REGION Network 25: STATE Num:70 StWtOTSFrmConv
   RUNG wire#powerrail
      Contact( #sStWtOTSFrmConv )
      wire#w1
      I_Contact( #sStWtResetRel )
      I_Contact( #sStWtOTSFrmConv_T1 )
      wire#w2
      Coil( #sStWtOTSFrmConv )
   END_RUNG
   RUNG wire#powerrail
      Contact( #sStWtL1S2DownOver_T1 )
   END_RUNG wire#w1
   RUNG wire#w2
      { S7_GenerateENO := "TRUE" } Move(in := 70, out1 => #StateNo)
   END_RUNG
   // the same network as SCL:
   #sStWtOTSFrmConv := (#sStWtOTSFrmConv OR #sStWtL1S2DownOver_T1) AND NOT #sStWtResetRel AND NOT #sStWtOTSFrmConv_T1;
   IF #sStWtOTSFrmConv THEN #StateNo := 70; END_IF;
END_REGION

REGION Network 26: Actions for STATE Num:70 StWtOTSFrmConv
   RUNG wire#powerrail
      Contact( #sStWtOTSFrmConv )
      Coil( #qRTRToConv )
   END_RUNG
   // the same network as SCL:
   #qRTRToConv := #sStWtOTSFrmConv;
END_REGION

REGION Network 27: Transition for STATE Num:80 StWtL1RecvBegin
   RUNG wire#powerrail
      Contact( #sStWtL1RecvBegin )
      I_Contact( #sStWtResetRel )
      Contact( #sSst )
      I_Contact( #iReceiveAreaClear )
      Coil( #sStWtL1RecvBegin_T1 )
   END_RUNG
   // the same network as SCL:
   #sStWtL1RecvBegin_T1 := #sStWtL1RecvBegin AND NOT #sStWtResetRel AND #sSst AND NOT #iReceiveAreaClear;
END_REGION

REGION Network 28: STATE Num:80 StWtL1RecvBegin
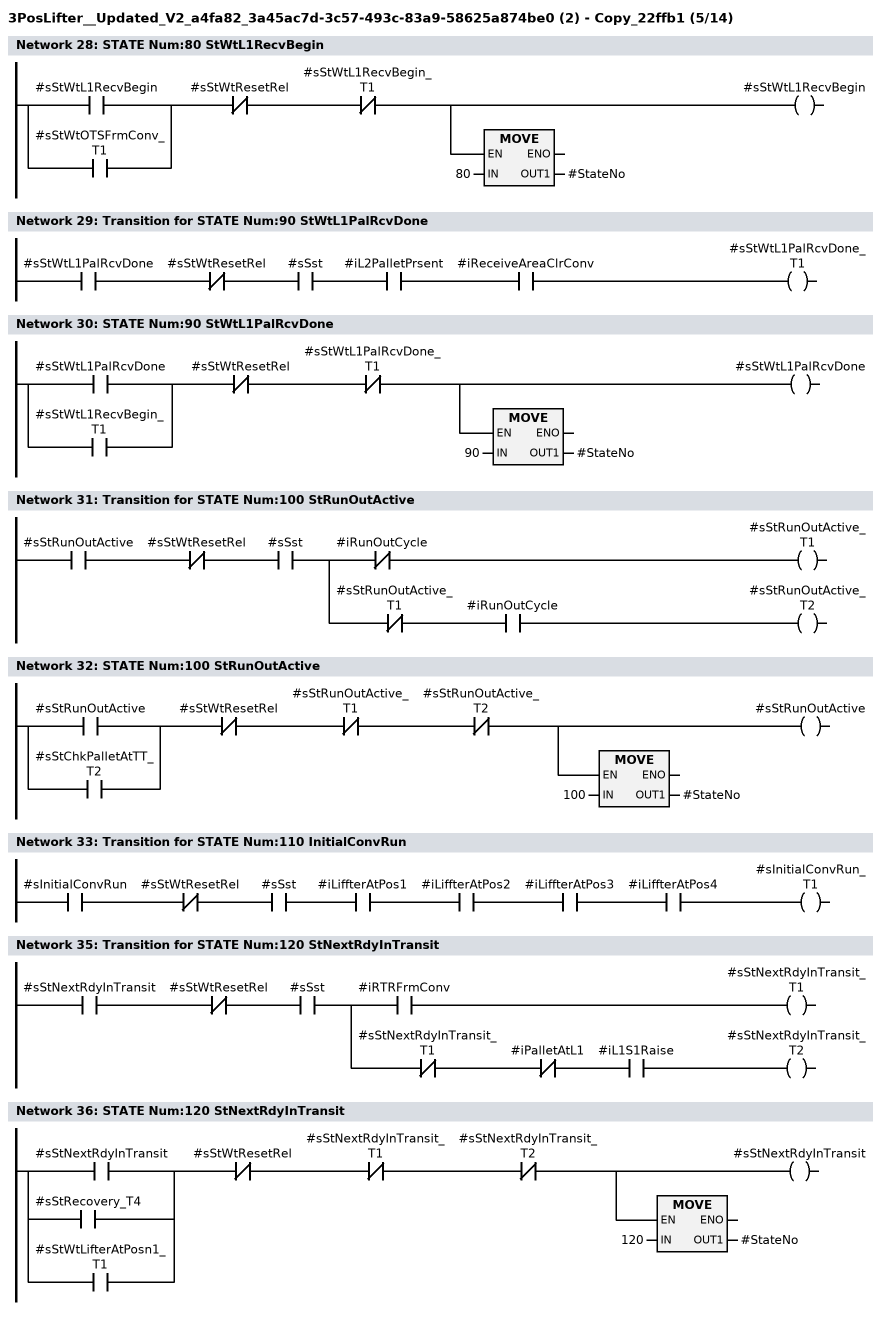
   RUNG wire#powerrail
      Contact( #sStWtL1RecvBegin )
      wire#w1
      I_Contact( #sStWtResetRel )
      I_Contact( #sStWtL1RecvBegin_T1 )
      wire#w2
      Coil( #sStWtL1RecvBegin )
   END_RUNG
   RUNG wire#powerrail
      Contact( #sStWtOTSFrmConv_T1 )
   END_RUNG wire#w1
   RUNG wire#w2
      { S7_GenerateENO := "TRUE" } Move(in := 80, out1 => #StateNo)
   END_RUNG
   // the same network as SCL:
   #sStWtL1RecvBegin := (#sStWtL1RecvBegin OR #sStWtOTSFrmConv_T1) AND NOT #sStWtResetRel AND NOT #sStWtL1RecvBegin_T1;
   IF #sStWtL1RecvBegin THEN #StateNo := 80; END_IF;
END_REGION

REGION Network 29: Transition for STATE Num:90 StWtL1PalRcvDone
   RUNG wire#powerrail
      Contact( #sStWtL1PalRcvDone )
      I_Contact( #sStWtResetRel )
      Contact( #sSst )
      Contact( #iL2PalletPrsent )
      Contact( #iReceiveAreaClrConv )
      Coil( #sStWtL1PalRcvDone_T1 )
   END_RUNG
   // the same network as SCL:
   #sStWtL1PalRcvDone_T1 := #sStWtL1PalRcvDone AND NOT #sStWtResetRel AND #sSst AND #iL2PalletPrsent AND #iReceiveAreaClrConv;
END_REGION

REGION Network 30: STATE Num:90 StWtL1PalRcvDone
   RUNG wire#powerrail
      Contact( #sStWtL1PalRcvDone )
      wire#w1
      I_Contact( #sStWtResetRel )
      I_Contact( #sStWtL1PalRcvDone_T1 )
      wire#w2
      Coil( #sStWtL1PalRcvDone )
   END_RUNG
   RUNG wire#powerrail
      Contact( #sStWtL1RecvBegin_T1 )
   END_RUNG wire#w1
   RUNG wire#w2
      { S7_GenerateENO := "TRUE" } Move(in := 90, out1 => #StateNo)
   END_RUNG
   // the same network as SCL:
   #sStWtL1PalRcvDone := (#sStWtL1PalRcvDone OR #sStWtL1RecvBegin_T1) AND NOT #sStWtResetRel AND NOT #sStWtL1PalRcvDone_T1;
   IF #sStWtL1PalRcvDone THEN #StateNo := 90; END_IF;
END_REGION

REGION Network 31: Transition for STATE Num:100 StRunOutActive
   RUNG wire#powerrail
      Contact( #sStRunOutActive )
      I_Contact( #sStWtResetRel )
      Contact( #sSst )
      wire#w1
      I_Contact( #iRunOutCycle )
      Coil( #sStRunOutActive_T1 )
   END_RUNG
   RUNG wire#w1
      I_Contact( #sStRunOutActive_T1 )
      Contact( #iRunOutCycle )
      Coil( #sStRunOutActive_T2 )
   END_RUNG
   // the same network as SCL:
   #_w1 := #sStRunOutActive AND NOT #sStWtResetRel AND #sSst;
   #sStRunOutActive_T1 := #_w1 AND NOT #iRunOutCycle;
   #sStRunOutActive_T2 := #_w1 AND NOT #sStRunOutActive_T1 AND #iRunOutCycle;
END_REGION

REGION Network 32: STATE Num:100 StRunOutActive
   RUNG wire#powerrail
      Contact( #sStRunOutActive )
      wire#w1
      I_Contact( #sStWtResetRel )
      I_Contact( #sStRunOutActive_T1 )
      I_Contact( #sStRunOutActive_T2 )
      wire#w2
      Coil( #sStRunOutActive )
   END_RUNG
   RUNG wire#powerrail
      Contact( #sStChkPalletAtTT_T2 )
   END_RUNG wire#w1
   RUNG wire#w2
      { S7_GenerateENO := "TRUE" } Move(in := 100, out1 => #StateNo)
   END_RUNG
   // the same network as SCL:
   #sStRunOutActive := (#sStRunOutActive OR #sStChkPalletAtTT_T2) AND NOT #sStWtResetRel AND NOT #sStRunOutActive_T1 AND NOT #sStRunOutActive_T2;
   IF #sStRunOutActive THEN #StateNo := 100; END_IF;
END_REGION

REGION Network 33: Transition for STATE Num:110 InitialConvRun
   RUNG wire#powerrail
      Contact( #sInitialConvRun )
      I_Contact( #sStWtResetRel )
      Contact( #sSst )
      Contact( #iLiffterAtPos1 )
      Contact( #iLiffterAtPos2 )
      Contact( #iLiffterAtPos3 )
      Contact( #iLiffterAtPos4 )
      Coil( #sInitialConvRun_T1 )
   END_RUNG
   // the same network as SCL:
   #sInitialConvRun_T1 := #sInitialConvRun AND NOT #sStWtResetRel AND #sSst AND #iLiffterAtPos1 AND #iLiffterAtPos2 AND #iLiffterAtPos3 AND #iLiffterAtPos4;
END_REGION

NETWORK
TITLE = STATE Num:110 InitialConvRun
      A(;
      O     #sInitialConvRun;
//wrong transition variable removed
      );
      AN    #sStWtResetRel;
      AN    #sInitialConvRun_T1;
      =     %L1.0;
      A     %L1.0;
      BLD   102;
      =     #sInitialConvRun;
      A     %L1.0;
      JNB   Label_110;
      L     110;
      T     #StateNo;
Label_110:NOP   0;

REGION Network 35: Transition for STATE Num:120 StNextRdyInTransit
   RUNG wire#powerrail
      Contact( #sStNextRdyInTransit )
      I_Contact( #sStWtResetRel )
      Contact( #sSst )
      wire#w1
      Contact( #iRTRFrmConv )
      Coil( #sStNextRdyInTransit_T1 )
   END_RUNG
   RUNG wire#w1
      I_Contact( #sStNextRdyInTransit_T1 )
      I_Contact( #iPalletAtL1 )
      Contact( #iL1S1Raise )
      Coil( #sStNextRdyInTransit_T2 )
   END_RUNG
   // the same network as SCL:
   #_w1 := #sStNextRdyInTransit AND NOT #sStWtResetRel AND #sSst;
   #sStNextRdyInTransit_T1 := #_w1 AND #iRTRFrmConv;
   #sStNextRdyInTransit_T2 := #_w1 AND NOT #sStNextRdyInTransit_T1 AND NOT #iPalletAtL1 AND #iL1S1Raise;
END_REGION

REGION Network 36: STATE Num:120 StNextRdyInTransit
   RUNG wire#powerrail
      Contact( #sStNextRdyInTransit )
      wire#w1
      I_Contact( #sStWtResetRel )
      I_Contact( #sStNextRdyInTransit_T1 )
      I_Contact( #sStNextRdyInTransit_T2 )
      wire#w2
      Coil( #sStNextRdyInTransit )
   END_RUNG
   RUNG wire#powerrail
      Contact( #sStRecovery_T4 )
   END_RUNG wire#w1
   RUNG wire#powerrail
      Contact( #sStWtLifterAtPosn1_T1 )
   END_RUNG wire#w1
   RUNG wire#w2
      { S7_GenerateENO := "TRUE" } Move(in := 120, out1 => #StateNo)
   END_RUNG
   // the same network as SCL:
   #sStNextRdyInTransit := (#sStNextRdyInTransit OR #sStRecovery_T4 OR #sStWtLifterAtPosn1_T1) AND NOT #sStWtResetRel AND NOT #sStNextRdyInTransit_T1 AND NOT #sStNextRdyInTransit_T2;
   IF #sStNextRdyInTransit THEN #StateNo := 120; END_IF;
END_REGION

REGION Network 37: Transition for STATE Num:130 StNextRdyInTransit_1
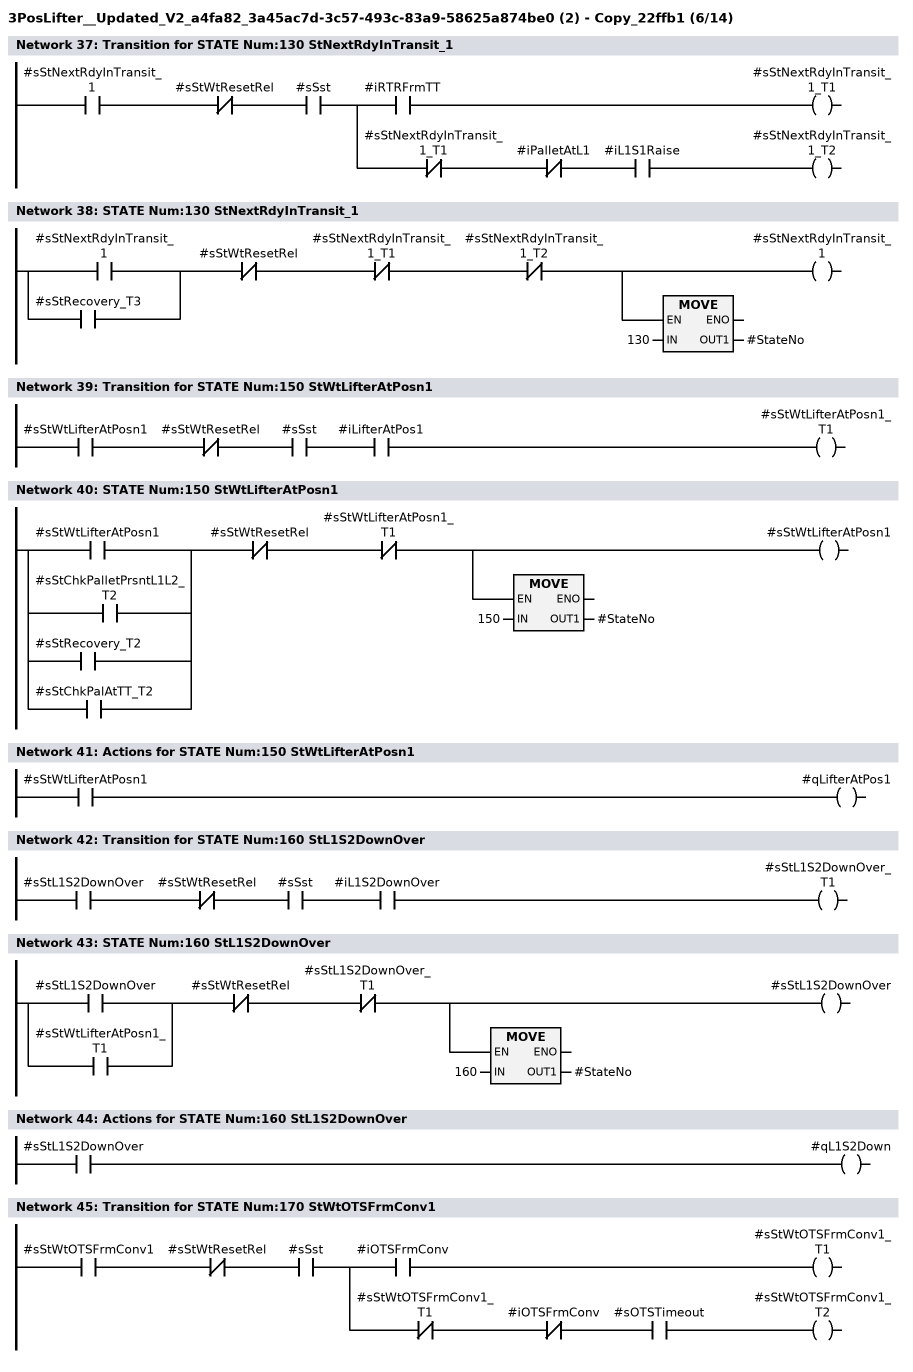
   RUNG wire#powerrail
      Contact( #sStNextRdyInTransit_1 )
      I_Contact( #sStWtResetRel )
      Contact( #sSst )
      wire#w1
      Contact( #iRTRFrmTT )
      Coil( #sStNextRdyInTransit_1_T1 )
   END_RUNG
   RUNG wire#w1
      I_Contact( #sStNextRdyInTransit_1_T1 )
      I_Contact( #iPalletAtL1 )
      Contact( #iL1S1Raise )
      Coil( #sStNextRdyInTransit_1_T2 )
   END_RUNG
   // the same network as SCL:
   #_w1 := #sStNextRdyInTransit_1 AND NOT #sStWtResetRel AND #sSst;
   #sStNextRdyInTransit_1_T1 := #_w1 AND #iRTRFrmTT;
   #sStNextRdyInTransit_1_T2 := #_w1 AND NOT #sStNextRdyInTransit_1_T1 AND NOT #iPalletAtL1 AND #iL1S1Raise;
END_REGION

REGION Network 38: STATE Num:130 StNextRdyInTransit_1
   RUNG wire#powerrail
      Contact( #sStNextRdyInTransit_1 )
      wire#w1
      I_Contact( #sStWtResetRel )
      I_Contact( #sStNextRdyInTransit_1_T1 )
      I_Contact( #sStNextRdyInTransit_1_T2 )
      wire#w2
      Coil( #sStNextRdyInTransit_1 )
   END_RUNG
   RUNG wire#powerrail
      Contact( #sStRecovery_T3 )
   END_RUNG wire#w1
   RUNG wire#w2
      { S7_GenerateENO := "TRUE" } Move(in := 130, out1 => #StateNo)
   END_RUNG
   // the same network as SCL:
   #sStNextRdyInTransit_1 := (#sStNextRdyInTransit_1 OR #sStRecovery_T3) AND NOT #sStWtResetRel AND NOT #sStNextRdyInTransit_1_T1 AND NOT #sStNextRdyInTransit_1_T2;
   IF #sStNextRdyInTransit_1 THEN #StateNo := 130; END_IF;
END_REGION

REGION Network 39: Transition for STATE Num:150 StWtLifterAtPosn1
   RUNG wire#powerrail
      Contact( #sStWtLifterAtPosn1 )
      I_Contact( #sStWtResetRel )
      Contact( #sSst )
      Contact( #iLifterAtPos1 )
      Coil( #sStWtLifterAtPosn1_T1 )
   END_RUNG
   // the same network as SCL:
   #sStWtLifterAtPosn1_T1 := #sStWtLifterAtPosn1 AND NOT #sStWtResetRel AND #sSst AND #iLifterAtPos1;
END_REGION

REGION Network 40: STATE Num:150 StWtLifterAtPosn1
   RUNG wire#powerrail
      Contact( #sStWtLifterAtPosn1 )
      wire#w1
      I_Contact( #sStWtResetRel )
      I_Contact( #sStWtLifterAtPosn1_T1 )
      wire#w2
      Coil( #sStWtLifterAtPosn1 )
   END_RUNG
   RUNG wire#powerrail
      Contact( #sStChkPalletPrsntL1L2_T2 )
   END_RUNG wire#w1
   RUNG wire#powerrail
      Contact( #sStRecovery_T2 )
   END_RUNG wire#w1
   RUNG wire#powerrail
      Contact( #sStChkPalAtTT_T2 )
   END_RUNG wire#w1
   RUNG wire#w2
      { S7_GenerateENO := "TRUE" } Move(in := 150, out1 => #StateNo)
   END_RUNG
   // the same network as SCL:
   #sStWtLifterAtPosn1 := (#sStWtLifterAtPosn1 OR #sStChkPalletPrsntL1L2_T2 OR #sStRecovery_T2 OR #sStChkPalAtTT_T2) AND NOT #sStWtResetRel AND NOT #sStWtLifterAtPosn1_T1;
   IF #sStWtLifterAtPosn1 THEN #StateNo := 150; END_IF;
END_REGION

REGION Network 41: Actions for STATE Num:150 StWtLifterAtPosn1
   RUNG wire#powerrail
      Contact( #sStWtLifterAtPosn1 )
      Coil( #qLifterAtPos1 )
   END_RUNG
   // the same network as SCL:
   #qLifterAtPos1 := #sStWtLifterAtPosn1;
END_REGION

REGION Network 42: Transition for STATE Num:160 StL1S2DownOver
   RUNG wire#powerrail
      Contact( #sStL1S2DownOver )
      I_Contact( #sStWtResetRel )
      Contact( #sSst )
      Contact( #iL1S2DownOver )
      Coil( #sStL1S2DownOver_T1 )
   END_RUNG
   // the same network as SCL:
   #sStL1S2DownOver_T1 := #sStL1S2DownOver AND NOT #sStWtResetRel AND #sSst AND #iL1S2DownOver;
END_REGION

REGION Network 43: STATE Num:160 StL1S2DownOver
   RUNG wire#powerrail
      Contact( #sStL1S2DownOver )
      wire#w1
      I_Contact( #sStWtResetRel )
      I_Contact( #sStL1S2DownOver_T1 )
      wire#w2
      Coil( #sStL1S2DownOver )
   END_RUNG
   RUNG wire#powerrail
      Contact( #sStWtLifterAtPosn1_T1 )
   END_RUNG wire#w1
   RUNG wire#w2
      { S7_GenerateENO := "TRUE" } Move(in := 160, out1 => #StateNo)
   END_RUNG
   // the same network as SCL:
   #sStL1S2DownOver := (#sStL1S2DownOver OR #sStWtLifterAtPosn1_T1) AND NOT #sStWtResetRel AND NOT #sStL1S2DownOver_T1;
   IF #sStL1S2DownOver THEN #StateNo := 160; END_IF;
END_REGION

REGION Network 44: Actions for STATE Num:160 StL1S2DownOver
   RUNG wire#powerrail
      Contact( #sStL1S2DownOver )
      Coil( #qL1S2Down )
   END_RUNG
   // the same network as SCL:
   #qL1S2Down := #sStL1S2DownOver;
END_REGION

REGION Network 45: Transition for STATE Num:170 StWtOTSFrmConv1
   RUNG wire#powerrail
      Contact( #sStWtOTSFrmConv1 )
      I_Contact( #sStWtResetRel )
      Contact( #sSst )
      wire#w1
      Contact( #iOTSFrmConv )
      Coil( #sStWtOTSFrmConv1_T1 )
   END_RUNG
   RUNG wire#w1
      I_Contact( #sStWtOTSFrmConv1_T1 )
      I_Contact( #iOTSFrmConv )
      Contact( #sOTSTimeout )
      Coil( #sStWtOTSFrmConv1_T2 )
   END_RUNG
   // the same network as SCL:
   #_w1 := #sStWtOTSFrmConv1 AND NOT #sStWtResetRel AND #sSst;
   #sStWtOTSFrmConv1_T1 := #_w1 AND #iOTSFrmConv;
   #sStWtOTSFrmConv1_T2 := #_w1 AND NOT #sStWtOTSFrmConv1_T1 AND NOT #iOTSFrmConv AND #sOTSTimeout;
END_REGION

REGION Network 46: STATE Num:170 StWtOTSFrmConv1
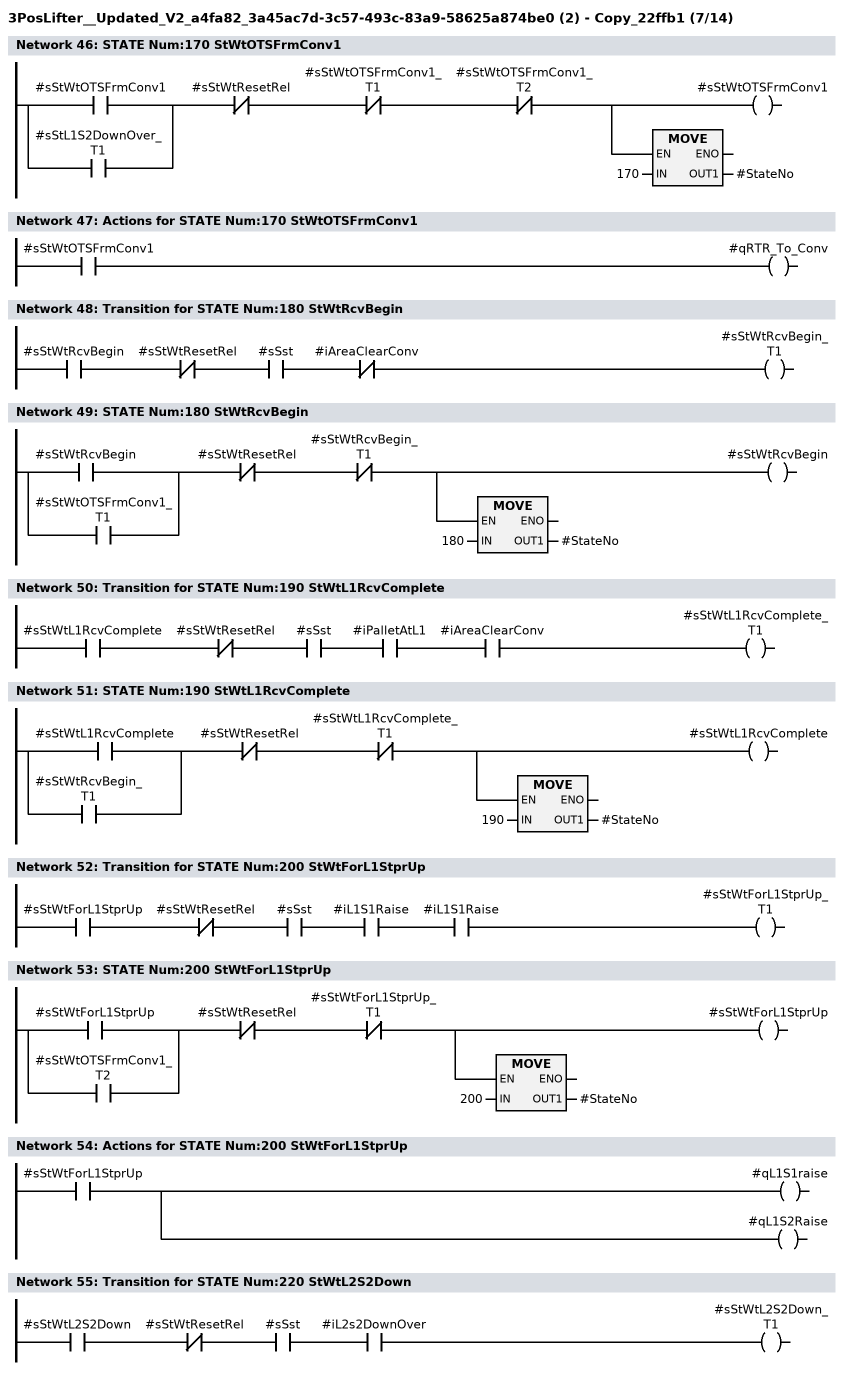
   RUNG wire#powerrail
      Contact( #sStWtOTSFrmConv1 )
      wire#w1
      I_Contact( #sStWtResetRel )
      I_Contact( #sStWtOTSFrmConv1_T1 )
      I_Contact( #sStWtOTSFrmConv1_T2 )
      wire#w2
      Coil( #sStWtOTSFrmConv1 )
   END_RUNG
   RUNG wire#powerrail
      Contact( #sStL1S2DownOver_T1 )
   END_RUNG wire#w1
   RUNG wire#w2
      { S7_GenerateENO := "TRUE" } Move(in := 170, out1 => #StateNo)
   END_RUNG
   // the same network as SCL:
   #sStWtOTSFrmConv1 := (#sStWtOTSFrmConv1 OR #sStL1S2DownOver_T1) AND NOT #sStWtResetRel AND NOT #sStWtOTSFrmConv1_T1 AND NOT #sStWtOTSFrmConv1_T2;
   IF #sStWtOTSFrmConv1 THEN #StateNo := 170; END_IF;
END_REGION

REGION Network 47: Actions for STATE Num:170 StWtOTSFrmConv1
   RUNG wire#powerrail
      Contact( #sStWtOTSFrmConv1 )
      Coil( #qRTR_To_Conv )
   END_RUNG
   // the same network as SCL:
   #qRTR_To_Conv := #sStWtOTSFrmConv1;
END_REGION

REGION Network 48: Transition for STATE Num:180 StWtRcvBegin
   RUNG wire#powerrail
      Contact( #sStWtRcvBegin )
      I_Contact( #sStWtResetRel )
      Contact( #sSst )
      I_Contact( #iAreaClearConv )
      Coil( #sStWtRcvBegin_T1 )
   END_RUNG
   // the same network as SCL:
   #sStWtRcvBegin_T1 := #sStWtRcvBegin AND NOT #sStWtResetRel AND #sSst AND NOT #iAreaClearConv;
END_REGION

REGION Network 49: STATE Num:180 StWtRcvBegin
   RUNG wire#powerrail
      Contact( #sStWtRcvBegin )
      wire#w1
      I_Contact( #sStWtResetRel )
      I_Contact( #sStWtRcvBegin_T1 )
      wire#w2
      Coil( #sStWtRcvBegin )
   END_RUNG
   RUNG wire#powerrail
      Contact( #sStWtOTSFrmConv1_T1 )
   END_RUNG wire#w1
   RUNG wire#w2
      { S7_GenerateENO := "TRUE" } Move(in := 180, out1 => #StateNo)
   END_RUNG
   // the same network as SCL:
   #sStWtRcvBegin := (#sStWtRcvBegin OR #sStWtOTSFrmConv1_T1) AND NOT #sStWtResetRel AND NOT #sStWtRcvBegin_T1;
   IF #sStWtRcvBegin THEN #StateNo := 180; END_IF;
END_REGION

REGION Network 50: Transition for STATE Num:190 StWtL1RcvComplete
   RUNG wire#powerrail
      Contact( #sStWtL1RcvComplete )
      I_Contact( #sStWtResetRel )
      Contact( #sSst )
      Contact( #iPalletAtL1 )
      Contact( #iAreaClearConv )
      Coil( #sStWtL1RcvComplete_T1 )
   END_RUNG
   // the same network as SCL:
   #sStWtL1RcvComplete_T1 := #sStWtL1RcvComplete AND NOT #sStWtResetRel AND #sSst AND #iPalletAtL1 AND #iAreaClearConv;
END_REGION

REGION Network 51: STATE Num:190 StWtL1RcvComplete
   RUNG wire#powerrail
      Contact( #sStWtL1RcvComplete )
      wire#w1
      I_Contact( #sStWtResetRel )
      I_Contact( #sStWtL1RcvComplete_T1 )
      wire#w2
      Coil( #sStWtL1RcvComplete )
   END_RUNG
   RUNG wire#powerrail
      Contact( #sStWtRcvBegin_T1 )
   END_RUNG wire#w1
   RUNG wire#w2
      { S7_GenerateENO := "TRUE" } Move(in := 190, out1 => #StateNo)
   END_RUNG
   // the same network as SCL:
   #sStWtL1RcvComplete := (#sStWtL1RcvComplete OR #sStWtRcvBegin_T1) AND NOT #sStWtResetRel AND NOT #sStWtL1RcvComplete_T1;
   IF #sStWtL1RcvComplete THEN #StateNo := 190; END_IF;
END_REGION

REGION Network 52: Transition for STATE Num:200 StWtForL1StprUp
   RUNG wire#powerrail
      Contact( #sStWtForL1StprUp )
      I_Contact( #sStWtResetRel )
      Contact( #sSst )
      Contact( #iL1S1Raise )
      Contact( #iL1S1Raise )
      Coil( #sStWtForL1StprUp_T1 )
   END_RUNG
   // the same network as SCL:
   #sStWtForL1StprUp_T1 := #sStWtForL1StprUp AND NOT #sStWtResetRel AND #sSst AND #iL1S1Raise AND #iL1S1Raise;
END_REGION

REGION Network 53: STATE Num:200 StWtForL1StprUp
   RUNG wire#powerrail
      Contact( #sStWtForL1StprUp )
      wire#w1
      I_Contact( #sStWtResetRel )
      I_Contact( #sStWtForL1StprUp_T1 )
      wire#w2
      Coil( #sStWtForL1StprUp )
   END_RUNG
   RUNG wire#powerrail
      Contact( #sStWtOTSFrmConv1_T2 )
   END_RUNG wire#w1
   RUNG wire#w2
      { S7_GenerateENO := "TRUE" } Move(in := 200, out1 => #StateNo)
   END_RUNG
   // the same network as SCL:
   #sStWtForL1StprUp := (#sStWtForL1StprUp OR #sStWtOTSFrmConv1_T2) AND NOT #sStWtResetRel AND NOT #sStWtForL1StprUp_T1;
   IF #sStWtForL1StprUp THEN #StateNo := 200; END_IF;
END_REGION

REGION Network 54: Actions for STATE Num:200 StWtForL1StprUp
   RUNG wire#powerrail
      Contact( #sStWtForL1StprUp )
      wire#w1
      Coil( #qL1S1raise )
   END_RUNG
   RUNG wire#w1
      Coil( #qL1S2Raise )
   END_RUNG
   // the same network as SCL:
   #qL1S1raise := #sStWtForL1StprUp;
   #qL1S2Raise := #sStWtForL1StprUp;
END_REGION

REGION Network 55: Transition for STATE Num:220 StWtL2S2Down
   RUNG wire#powerrail
      Contact( #sStWtL2S2Down )
      I_Contact( #sStWtResetRel )
      Contact( #sSst )
      Contact( #iL2s2DownOver )
      Coil( #sStWtL2S2Down_T1 )
   END_RUNG
   // the same network as SCL:
   #sStWtL2S2Down_T1 := #sStWtL2S2Down AND NOT #sStWtResetRel AND #sSst AND #iL2s2DownOver;
END_REGION

REGION Network 56: STATE Num:220 StWtL2S2Down
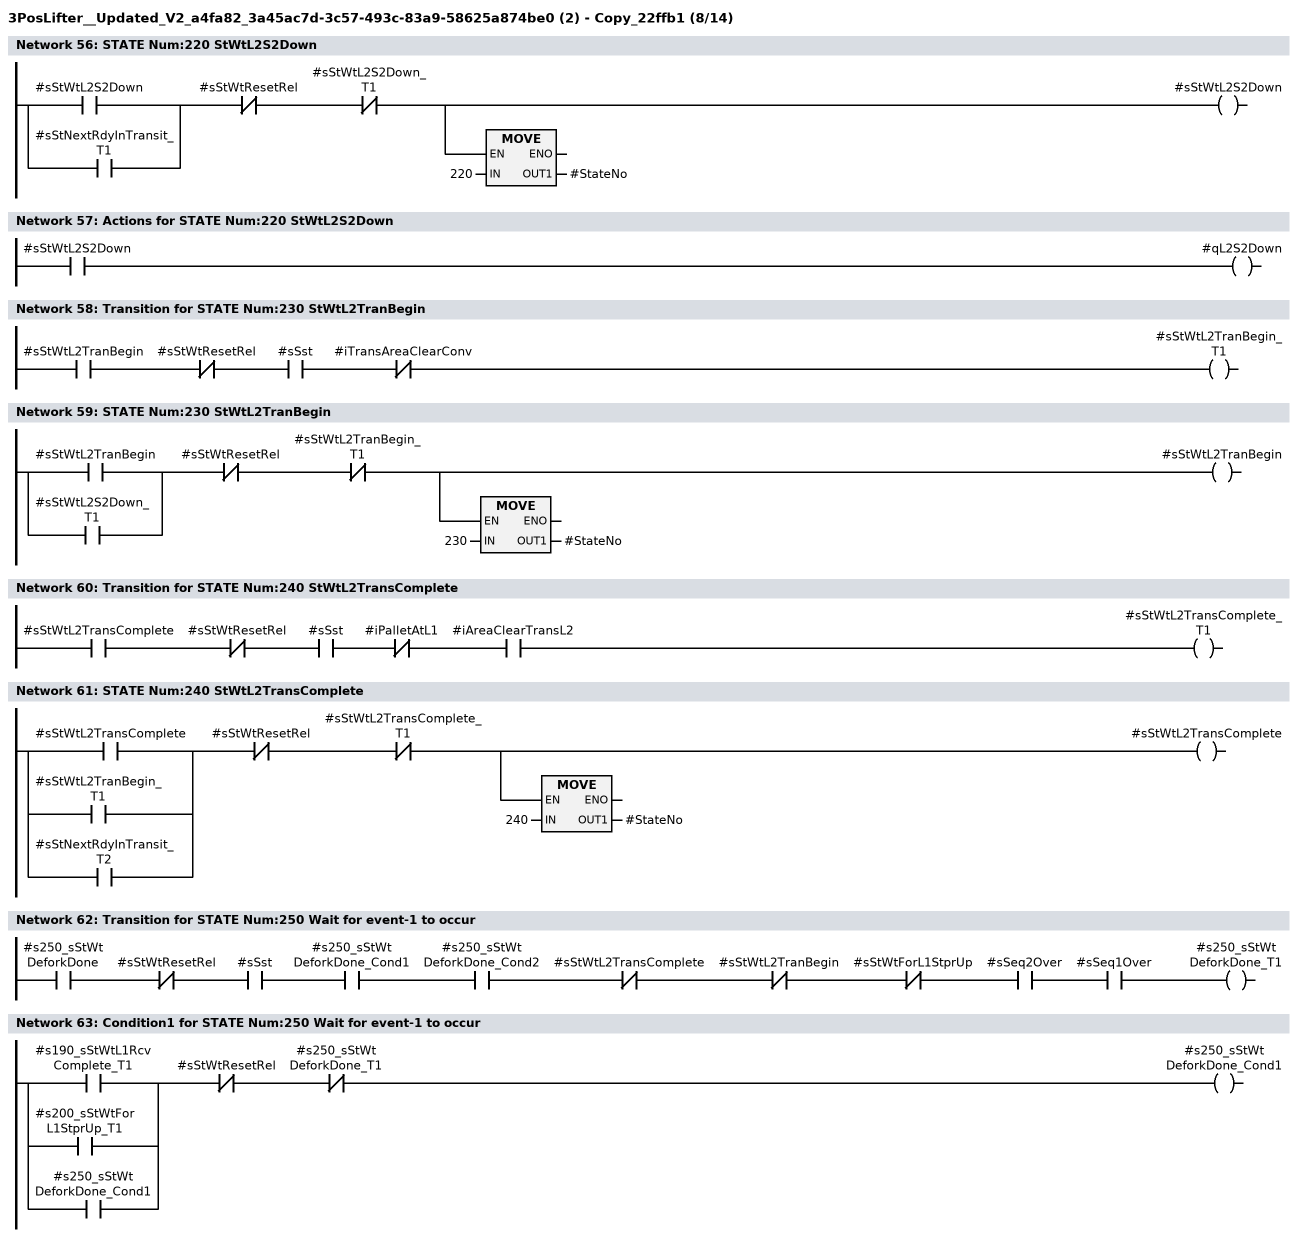
   RUNG wire#powerrail
      Contact( #sStWtL2S2Down )
      wire#w1
      I_Contact( #sStWtResetRel )
      I_Contact( #sStWtL2S2Down_T1 )
      wire#w2
      Coil( #sStWtL2S2Down )
   END_RUNG
   RUNG wire#powerrail
      Contact( #sStNextRdyInTransit_T1 )
   END_RUNG wire#w1
   RUNG wire#w2
      { S7_GenerateENO := "TRUE" } Move(in := 220, out1 => #StateNo)
   END_RUNG
   // the same network as SCL:
   #sStWtL2S2Down := (#sStWtL2S2Down OR #sStNextRdyInTransit_T1) AND NOT #sStWtResetRel AND NOT #sStWtL2S2Down_T1;
   IF #sStWtL2S2Down THEN #StateNo := 220; END_IF;
END_REGION

REGION Network 57: Actions for STATE Num:220 StWtL2S2Down
   RUNG wire#powerrail
      Contact( #sStWtL2S2Down )
      Coil( #qL2S2Down )
   END_RUNG
   // the same network as SCL:
   #qL2S2Down := #sStWtL2S2Down;
END_REGION

REGION Network 58: Transition for STATE Num:230 StWtL2TranBegin
   RUNG wire#powerrail
      Contact( #sStWtL2TranBegin )
      I_Contact( #sStWtResetRel )
      Contact( #sSst )
      I_Contact( #iTransAreaClearConv )
      Coil( #sStWtL2TranBegin_T1 )
   END_RUNG
   // the same network as SCL:
   #sStWtL2TranBegin_T1 := #sStWtL2TranBegin AND NOT #sStWtResetRel AND #sSst AND NOT #iTransAreaClearConv;
END_REGION

REGION Network 59: STATE Num:230 StWtL2TranBegin
   RUNG wire#powerrail
      Contact( #sStWtL2TranBegin )
      wire#w1
      I_Contact( #sStWtResetRel )
      I_Contact( #sStWtL2TranBegin_T1 )
      wire#w2
      Coil( #sStWtL2TranBegin )
   END_RUNG
   RUNG wire#powerrail
      Contact( #sStWtL2S2Down_T1 )
   END_RUNG wire#w1
   RUNG wire#w2
      { S7_GenerateENO := "TRUE" } Move(in := 230, out1 => #StateNo)
   END_RUNG
   // the same network as SCL:
   #sStWtL2TranBegin := (#sStWtL2TranBegin OR #sStWtL2S2Down_T1) AND NOT #sStWtResetRel AND NOT #sStWtL2TranBegin_T1;
   IF #sStWtL2TranBegin THEN #StateNo := 230; END_IF;
END_REGION

REGION Network 60: Transition for STATE Num:240 StWtL2TransComplete
   RUNG wire#powerrail
      Contact( #sStWtL2TransComplete )
      I_Contact( #sStWtResetRel )
      Contact( #sSst )
      I_Contact( #iPalletAtL1 )
      Contact( #iAreaClearTransL2 )
      Coil( #sStWtL2TransComplete_T1 )
   END_RUNG
   // the same network as SCL:
   #sStWtL2TransComplete_T1 := #sStWtL2TransComplete AND NOT #sStWtResetRel AND #sSst AND NOT #iPalletAtL1 AND #iAreaClearTransL2;
END_REGION

REGION Network 61: STATE Num:240 StWtL2TransComplete
   RUNG wire#powerrail
      Contact( #sStWtL2TransComplete )
      wire#w1
      I_Contact( #sStWtResetRel )
      I_Contact( #sStWtL2TransComplete_T1 )
      wire#w2
      Coil( #sStWtL2TransComplete )
   END_RUNG
   RUNG wire#powerrail
      Contact( #sStWtL2TranBegin_T1 )
   END_RUNG wire#w1
   RUNG wire#powerrail
      Contact( #sStNextRdyInTransit_T2 )
   END_RUNG wire#w1
   RUNG wire#w2
      { S7_GenerateENO := "TRUE" } Move(in := 240, out1 => #StateNo)
   END_RUNG
   // the same network as SCL:
   #sStWtL2TransComplete := (#sStWtL2TransComplete OR #sStWtL2TranBegin_T1 OR #sStNextRdyInTransit_T2) AND NOT #sStWtResetRel AND NOT #sStWtL2TransComplete_T1;
   IF #sStWtL2TransComplete THEN #StateNo := 240; END_IF;
END_REGION

REGION Network 62: Transition for STATE Num:250 Wait for event-1 to occur
   RUNG wire#powerrail
      Contact( #s250_sStWtDeforkDone )
      I_Contact( #sStWtResetRel )
      Contact( #sSst )
      Contact( #s250_sStWtDeforkDone_Cond1 )
      Contact( #s250_sStWtDeforkDone_Cond2 )
      I_Contact( #sStWtL2TransComplete )
      I_Contact( #sStWtL2TranBegin )
      I_Contact( #sStWtForL1StprUp )
      Contact( #sSeq2Over )
      Contact( #sSeq1Over )
      Coil( #s250_sStWtDeforkDone_T1 )
   END_RUNG
   // the same network as SCL:
   #s250_sStWtDeforkDone_T1 := #s250_sStWtDeforkDone AND NOT #sStWtResetRel AND #sSst AND #s250_sStWtDeforkDone_Cond1 AND #s250_sStWtDeforkDone_Cond2 AND NOT #sStWtL2TransComplete AND NOT #sStWtL2TranBegin AND NOT #sStWtForL1StprUp AND #sSeq2Over AND #sSeq1Over;
END_REGION

REGION Network 63: Condition1 for STATE Num:250 Wait for event-1 to occur
   RUNG wire#powerrail
      Contact( #s190_sStWtL1RcvComplete_T1 )
      wire#w1
      I_Contact( #sStWtResetRel )
      I_Contact( #s250_sStWtDeforkDone_T1 )
      Coil( #s250_sStWtDeforkDone_Cond1 )
   END_RUNG
   RUNG wire#powerrail
      Contact( #s200_sStWtForL1StprUp_T1 )
   END_RUNG wire#w1
   RUNG wire#powerrail
      Contact( #s250_sStWtDeforkDone_Cond1 )
   END_RUNG wire#w1
   // the same network as SCL:
   #s250_sStWtDeforkDone_Cond1 := (#s190_sStWtL1RcvComplete_T1 OR #s200_sStWtForL1StprUp_T1 OR #s250_sStWtDeforkDone_Cond1) AND NOT #sStWtResetRel AND NOT #s250_sStWtDeforkDone_T1;
END_REGION

REGION Network 64: Condition2 for STATE Num:250 Wait for event-1 to occur
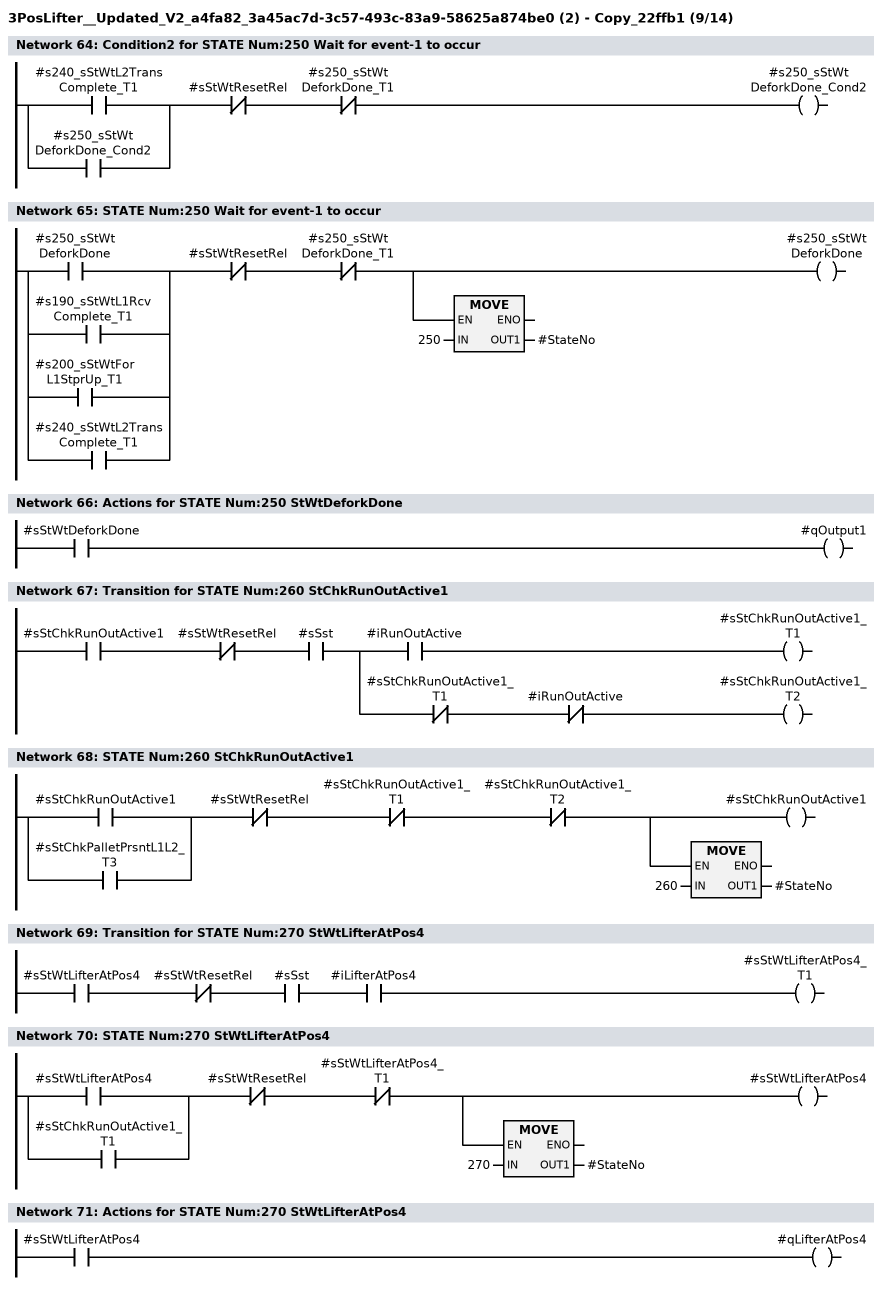
   RUNG wire#powerrail
      Contact( #s240_sStWtL2TransComplete_T1 )
      wire#w1
      I_Contact( #sStWtResetRel )
      I_Contact( #s250_sStWtDeforkDone_T1 )
      Coil( #s250_sStWtDeforkDone_Cond2 )
   END_RUNG
   RUNG wire#powerrail
      Contact( #s250_sStWtDeforkDone_Cond2 )
   END_RUNG wire#w1
   // the same network as SCL:
   #s250_sStWtDeforkDone_Cond2 := (#s240_sStWtL2TransComplete_T1 OR #s250_sStWtDeforkDone_Cond2) AND NOT #sStWtResetRel AND NOT #s250_sStWtDeforkDone_T1;
END_REGION

REGION Network 65: STATE Num:250 Wait for event-1 to occur
   RUNG wire#powerrail
      Contact( #s250_sStWtDeforkDone )
      wire#w1
      I_Contact( #sStWtResetRel )
      I_Contact( #s250_sStWtDeforkDone_T1 )
      wire#w2
      Coil( #s250_sStWtDeforkDone )
   END_RUNG
   RUNG wire#powerrail
      Contact( #s190_sStWtL1RcvComplete_T1 )
   END_RUNG wire#w1
   RUNG wire#powerrail
      Contact( #s200_sStWtForL1StprUp_T1 )
   END_RUNG wire#w1
   RUNG wire#powerrail
      Contact( #s240_sStWtL2TransComplete_T1 )
   END_RUNG wire#w1
   RUNG wire#w2
      { S7_GenerateENO := "TRUE" } Move(in := 250, out1 => #StateNo)
   END_RUNG
   // the same network as SCL:
   #s250_sStWtDeforkDone := (#s250_sStWtDeforkDone OR #s190_sStWtL1RcvComplete_T1 OR #s200_sStWtForL1StprUp_T1 OR #s240_sStWtL2TransComplete_T1) AND NOT #sStWtResetRel AND NOT #s250_sStWtDeforkDone_T1;
   IF #s250_sStWtDeforkDone THEN #StateNo := 250; END_IF;
END_REGION

REGION Network 66: Actions for STATE Num:250 StWtDeforkDone
   RUNG wire#powerrail
      Contact( #sStWtDeforkDone )
      Coil( #qOutput1 )
   END_RUNG
   // the same network as SCL:
   #qOutput1 := #sStWtDeforkDone;
END_REGION

REGION Network 67: Transition for STATE Num:260 StChkRunOutActive1
   RUNG wire#powerrail
      Contact( #sStChkRunOutActive1 )
      I_Contact( #sStWtResetRel )
      Contact( #sSst )
      wire#w1
      Contact( #iRunOutActive )
      Coil( #sStChkRunOutActive1_T1 )
   END_RUNG
   RUNG wire#w1
      I_Contact( #sStChkRunOutActive1_T1 )
      I_Contact( #iRunOutActive )
      Coil( #sStChkRunOutActive1_T2 )
   END_RUNG
   // the same network as SCL:
   #_w1 := #sStChkRunOutActive1 AND NOT #sStWtResetRel AND #sSst;
   #sStChkRunOutActive1_T1 := #_w1 AND #iRunOutActive;
   #sStChkRunOutActive1_T2 := #_w1 AND NOT #sStChkRunOutActive1_T1 AND NOT #iRunOutActive;
END_REGION

REGION Network 68: STATE Num:260 StChkRunOutActive1
   RUNG wire#powerrail
      Contact( #sStChkRunOutActive1 )
      wire#w1
      I_Contact( #sStWtResetRel )
      I_Contact( #sStChkRunOutActive1_T1 )
      I_Contact( #sStChkRunOutActive1_T2 )
      wire#w2
      Coil( #sStChkRunOutActive1 )
   END_RUNG
   RUNG wire#powerrail
      Contact( #sStChkPalletPrsntL1L2_T3 )
   END_RUNG wire#w1
   RUNG wire#w2
      { S7_GenerateENO := "TRUE" } Move(in := 260, out1 => #StateNo)
   END_RUNG
   // the same network as SCL:
   #sStChkRunOutActive1 := (#sStChkRunOutActive1 OR #sStChkPalletPrsntL1L2_T3) AND NOT #sStWtResetRel AND NOT #sStChkRunOutActive1_T1 AND NOT #sStChkRunOutActive1_T2;
   IF #sStChkRunOutActive1 THEN #StateNo := 260; END_IF;
END_REGION

REGION Network 69: Transition for STATE Num:270 StWtLifterAtPos4
   RUNG wire#powerrail
      Contact( #sStWtLifterAtPos4 )
      I_Contact( #sStWtResetRel )
      Contact( #sSst )
      Contact( #iLifterAtPos4 )
      Coil( #sStWtLifterAtPos4_T1 )
   END_RUNG
   // the same network as SCL:
   #sStWtLifterAtPos4_T1 := #sStWtLifterAtPos4 AND NOT #sStWtResetRel AND #sSst AND #iLifterAtPos4;
END_REGION

REGION Network 70: STATE Num:270 StWtLifterAtPos4
   RUNG wire#powerrail
      Contact( #sStWtLifterAtPos4 )
      wire#w1
      I_Contact( #sStWtResetRel )
      I_Contact( #sStWtLifterAtPos4_T1 )
      wire#w2
      Coil( #sStWtLifterAtPos4 )
   END_RUNG
   RUNG wire#powerrail
      Contact( #sStChkRunOutActive1_T1 )
   END_RUNG wire#w1
   RUNG wire#w2
      { S7_GenerateENO := "TRUE" } Move(in := 270, out1 => #StateNo)
   END_RUNG
   // the same network as SCL:
   #sStWtLifterAtPos4 := (#sStWtLifterAtPos4 OR #sStChkRunOutActive1_T1) AND NOT #sStWtResetRel AND NOT #sStWtLifterAtPos4_T1;
   IF #sStWtLifterAtPos4 THEN #StateNo := 270; END_IF;
END_REGION

REGION Network 71: Actions for STATE Num:270 StWtLifterAtPos4
   RUNG wire#powerrail
      Contact( #sStWtLifterAtPos4 )
      Coil( #qLifterAtPos4 )
   END_RUNG
   // the same network as SCL:
   #qLifterAtPos4 := #sStWtLifterAtPos4;
END_REGION

REGION Network 72: Transition for STATE Num:280 StWtRTRFrmConvPos4
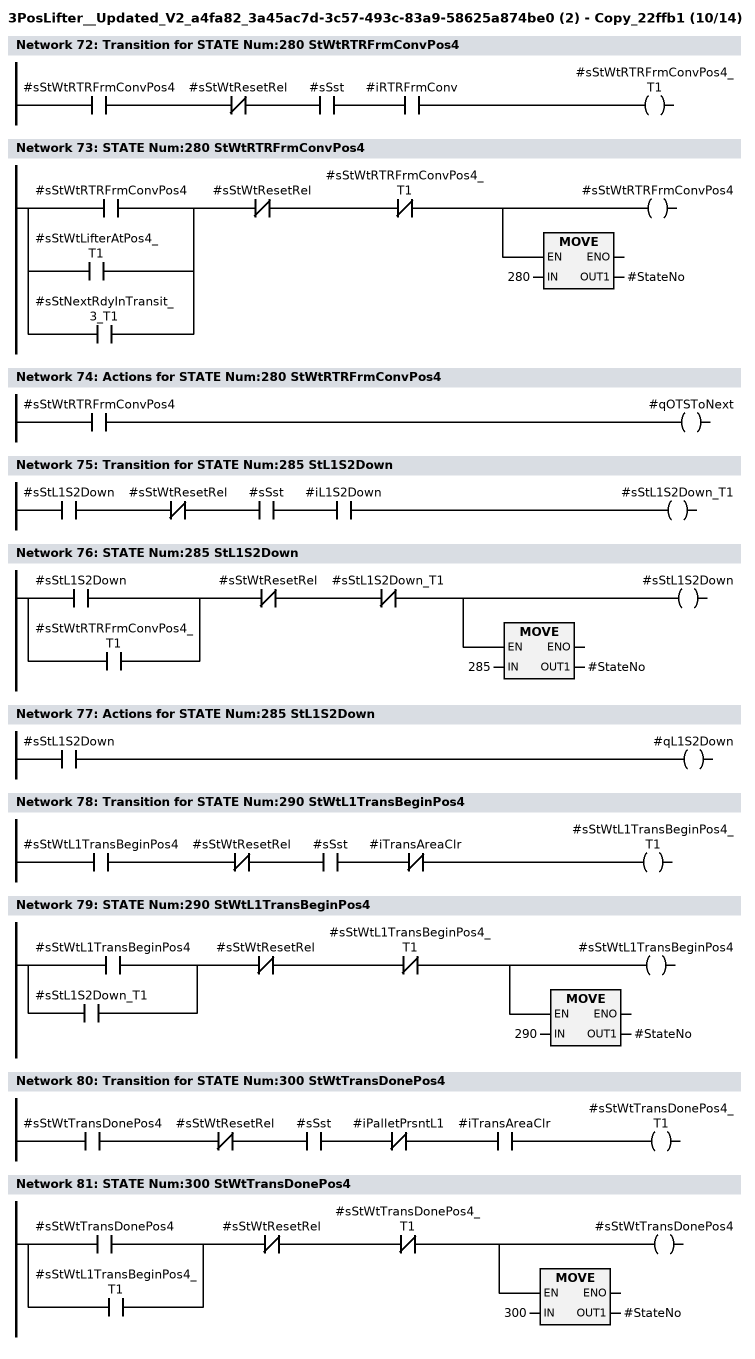
   RUNG wire#powerrail
      Contact( #sStWtRTRFrmConvPos4 )
      I_Contact( #sStWtResetRel )
      Contact( #sSst )
      Contact( #iRTRFrmConv )
      Coil( #sStWtRTRFrmConvPos4_T1 )
   END_RUNG
   // the same network as SCL:
   #sStWtRTRFrmConvPos4_T1 := #sStWtRTRFrmConvPos4 AND NOT #sStWtResetRel AND #sSst AND #iRTRFrmConv;
END_REGION

REGION Network 73: STATE Num:280 StWtRTRFrmConvPos4
   RUNG wire#powerrail
      Contact( #sStWtRTRFrmConvPos4 )
      wire#w1
      I_Contact( #sStWtResetRel )
      I_Contact( #sStWtRTRFrmConvPos4_T1 )
      wire#w2
      Coil( #sStWtRTRFrmConvPos4 )
   END_RUNG
   RUNG wire#powerrail
      Contact( #sStWtLifterAtPos4_T1 )
   END_RUNG wire#w1
   RUNG wire#powerrail
      Contact( #sStNextRdyInTransit_3_T1 )
   END_RUNG wire#w1
   RUNG wire#w2
      { S7_GenerateENO := "TRUE" } Move(in := 280, out1 => #StateNo)
   END_RUNG
   // the same network as SCL:
   #sStWtRTRFrmConvPos4 := (#sStWtRTRFrmConvPos4 OR #sStWtLifterAtPos4_T1 OR #sStNextRdyInTransit_3_T1) AND NOT #sStWtResetRel AND NOT #sStWtRTRFrmConvPos4_T1;
   IF #sStWtRTRFrmConvPos4 THEN #StateNo := 280; END_IF;
END_REGION

REGION Network 74: Actions for STATE Num:280 StWtRTRFrmConvPos4
   RUNG wire#powerrail
      Contact( #sStWtRTRFrmConvPos4 )
      Coil( #qOTSToNext )
   END_RUNG
   // the same network as SCL:
   #qOTSToNext := #sStWtRTRFrmConvPos4;
END_REGION

REGION Network 75: Transition for STATE Num:285 StL1S2Down
   RUNG wire#powerrail
      Contact( #sStL1S2Down )
      I_Contact( #sStWtResetRel )
      Contact( #sSst )
      Contact( #iL1S2Down )
      Coil( #sStL1S2Down_T1 )
   END_RUNG
   // the same network as SCL:
   #sStL1S2Down_T1 := #sStL1S2Down AND NOT #sStWtResetRel AND #sSst AND #iL1S2Down;
END_REGION

REGION Network 76: STATE Num:285 StL1S2Down
   RUNG wire#powerrail
      Contact( #sStL1S2Down )
      wire#w1
      I_Contact( #sStWtResetRel )
      I_Contact( #sStL1S2Down_T1 )
      wire#w2
      Coil( #sStL1S2Down )
   END_RUNG
   RUNG wire#powerrail
      Contact( #sStWtRTRFrmConvPos4_T1 )
   END_RUNG wire#w1
   RUNG wire#w2
      { S7_GenerateENO := "TRUE" } Move(in := 285, out1 => #StateNo)
   END_RUNG
   // the same network as SCL:
   #sStL1S2Down := (#sStL1S2Down OR #sStWtRTRFrmConvPos4_T1) AND NOT #sStWtResetRel AND NOT #sStL1S2Down_T1;
   IF #sStL1S2Down THEN #StateNo := 285; END_IF;
END_REGION

REGION Network 77: Actions for STATE Num:285 StL1S2Down
   RUNG wire#powerrail
      Contact( #sStL1S2Down )
      Coil( #qL1S2Down )
   END_RUNG
   // the same network as SCL:
   #qL1S2Down := #sStL1S2Down;
END_REGION

REGION Network 78: Transition for STATE Num:290 StWtL1TransBeginPos4
   RUNG wire#powerrail
      Contact( #sStWtL1TransBeginPos4 )
      I_Contact( #sStWtResetRel )
      Contact( #sSst )
      I_Contact( #iTransAreaClr )
      Coil( #sStWtL1TransBeginPos4_T1 )
   END_RUNG
   // the same network as SCL:
   #sStWtL1TransBeginPos4_T1 := #sStWtL1TransBeginPos4 AND NOT #sStWtResetRel AND #sSst AND NOT #iTransAreaClr;
END_REGION

REGION Network 79: STATE Num:290 StWtL1TransBeginPos4
   RUNG wire#powerrail
      Contact( #sStWtL1TransBeginPos4 )
      wire#w1
      I_Contact( #sStWtResetRel )
      I_Contact( #sStWtL1TransBeginPos4_T1 )
      wire#w2
      Coil( #sStWtL1TransBeginPos4 )
   END_RUNG
   RUNG wire#powerrail
      Contact( #sStL1S2Down_T1 )
   END_RUNG wire#w1
   RUNG wire#w2
      { S7_GenerateENO := "TRUE" } Move(in := 290, out1 => #StateNo)
   END_RUNG
   // the same network as SCL:
   #sStWtL1TransBeginPos4 := (#sStWtL1TransBeginPos4 OR #sStL1S2Down_T1) AND NOT #sStWtResetRel AND NOT #sStWtL1TransBeginPos4_T1;
   IF #sStWtL1TransBeginPos4 THEN #StateNo := 290; END_IF;
END_REGION

REGION Network 80: Transition for STATE Num:300 StWtTransDonePos4
   RUNG wire#powerrail
      Contact( #sStWtTransDonePos4 )
      I_Contact( #sStWtResetRel )
      Contact( #sSst )
      I_Contact( #iPalletPrsntL1 )
      Contact( #iTransAreaClr )
      Coil( #sStWtTransDonePos4_T1 )
   END_RUNG
   // the same network as SCL:
   #sStWtTransDonePos4_T1 := #sStWtTransDonePos4 AND NOT #sStWtResetRel AND #sSst AND NOT #iPalletPrsntL1 AND #iTransAreaClr;
END_REGION

REGION Network 81: STATE Num:300 StWtTransDonePos4
   RUNG wire#powerrail
      Contact( #sStWtTransDonePos4 )
      wire#w1
      I_Contact( #sStWtResetRel )
      I_Contact( #sStWtTransDonePos4_T1 )
      wire#w2
      Coil( #sStWtTransDonePos4 )
   END_RUNG
   RUNG wire#powerrail
      Contact( #sStWtL1TransBeginPos4_T1 )
   END_RUNG wire#w1
   RUNG wire#w2
      { S7_GenerateENO := "TRUE" } Move(in := 300, out1 => #StateNo)
   END_RUNG
   // the same network as SCL:
   #sStWtTransDonePos4 := (#sStWtTransDonePos4 OR #sStWtL1TransBeginPos4_T1) AND NOT #sStWtResetRel AND NOT #sStWtTransDonePos4_T1;
   IF #sStWtTransDonePos4 THEN #StateNo := 300; END_IF;
END_REGION

REGION Network 82: Transition for STATE Num:310 StChkPalletAtTT1
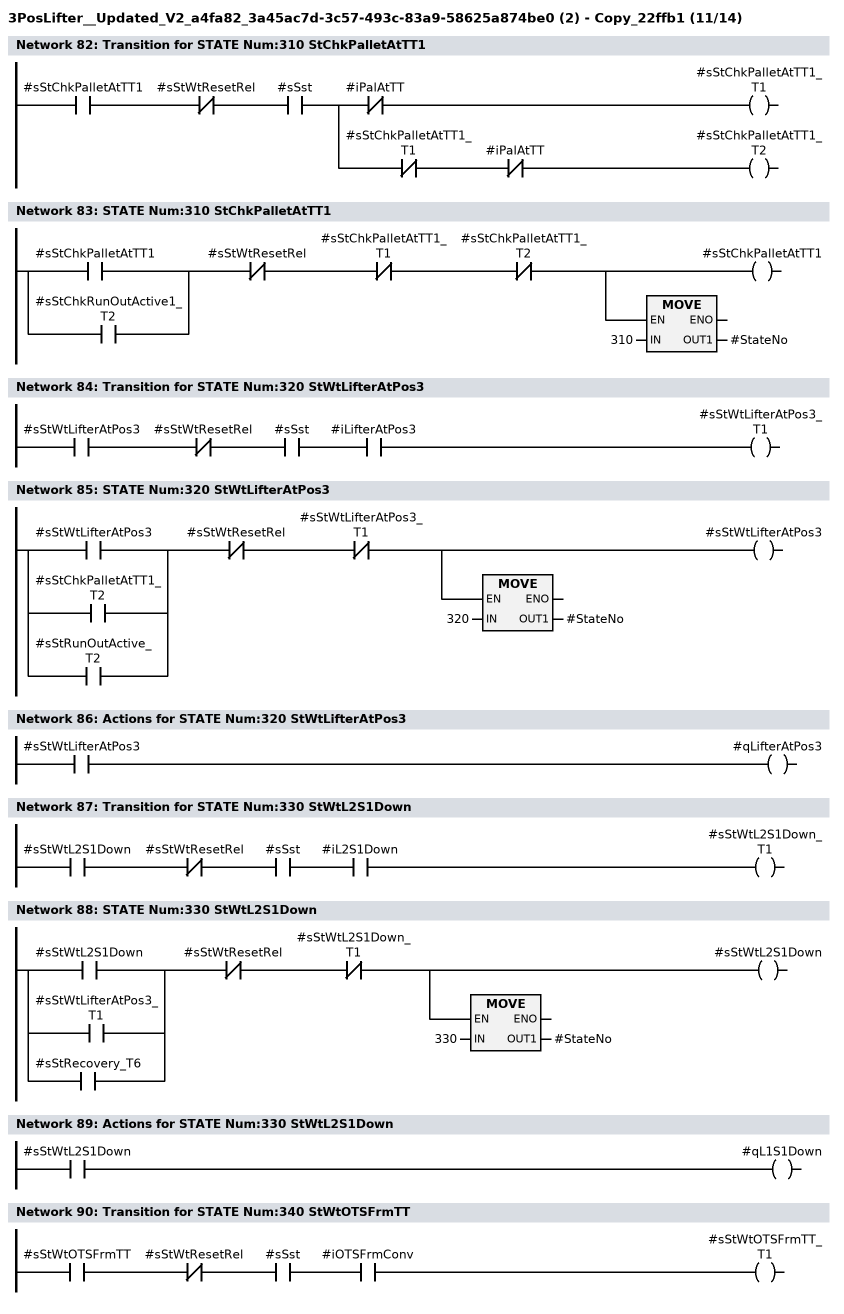
   RUNG wire#powerrail
      Contact( #sStChkPalletAtTT1 )
      I_Contact( #sStWtResetRel )
      Contact( #sSst )
      wire#w1
      I_Contact( #iPalAtTT )
      Coil( #sStChkPalletAtTT1_T1 )
   END_RUNG
   RUNG wire#w1
      I_Contact( #sStChkPalletAtTT1_T1 )
      I_Contact( #iPalAtTT )
      Coil( #sStChkPalletAtTT1_T2 )
   END_RUNG
   // the same network as SCL:
   #_w1 := #sStChkPalletAtTT1 AND NOT #sStWtResetRel AND #sSst;
   #sStChkPalletAtTT1_T1 := #_w1 AND NOT #iPalAtTT;
   #sStChkPalletAtTT1_T2 := #_w1 AND NOT #sStChkPalletAtTT1_T1 AND NOT #iPalAtTT;
END_REGION

REGION Network 83: STATE Num:310 StChkPalletAtTT1
   RUNG wire#powerrail
      Contact( #sStChkPalletAtTT1 )
      wire#w1
      I_Contact( #sStWtResetRel )
      I_Contact( #sStChkPalletAtTT1_T1 )
      I_Contact( #sStChkPalletAtTT1_T2 )
      wire#w2
      Coil( #sStChkPalletAtTT1 )
   END_RUNG
   RUNG wire#powerrail
      Contact( #sStChkRunOutActive1_T2 )
   END_RUNG wire#w1
   RUNG wire#w2
      { S7_GenerateENO := "TRUE" } Move(in := 310, out1 => #StateNo)
   END_RUNG
   // the same network as SCL:
   #sStChkPalletAtTT1 := (#sStChkPalletAtTT1 OR #sStChkRunOutActive1_T2) AND NOT #sStWtResetRel AND NOT #sStChkPalletAtTT1_T1 AND NOT #sStChkPalletAtTT1_T2;
   IF #sStChkPalletAtTT1 THEN #StateNo := 310; END_IF;
END_REGION

REGION Network 84: Transition for STATE Num:320 StWtLifterAtPos3
   RUNG wire#powerrail
      Contact( #sStWtLifterAtPos3 )
      I_Contact( #sStWtResetRel )
      Contact( #sSst )
      Contact( #iLifterAtPos3 )
      Coil( #sStWtLifterAtPos3_T1 )
   END_RUNG
   // the same network as SCL:
   #sStWtLifterAtPos3_T1 := #sStWtLifterAtPos3 AND NOT #sStWtResetRel AND #sSst AND #iLifterAtPos3;
END_REGION

REGION Network 85: STATE Num:320 StWtLifterAtPos3
   RUNG wire#powerrail
      Contact( #sStWtLifterAtPos3 )
      wire#w1
      I_Contact( #sStWtResetRel )
      I_Contact( #sStWtLifterAtPos3_T1 )
      wire#w2
      Coil( #sStWtLifterAtPos3 )
   END_RUNG
   RUNG wire#powerrail
      Contact( #sStChkPalletAtTT1_T2 )
   END_RUNG wire#w1
   RUNG wire#powerrail
      Contact( #sStRunOutActive_T2 )
   END_RUNG wire#w1
   RUNG wire#w2
      { S7_GenerateENO := "TRUE" } Move(in := 320, out1 => #StateNo)
   END_RUNG
   // the same network as SCL:
   #sStWtLifterAtPos3 := (#sStWtLifterAtPos3 OR #sStChkPalletAtTT1_T2 OR #sStRunOutActive_T2) AND NOT #sStWtResetRel AND NOT #sStWtLifterAtPos3_T1;
   IF #sStWtLifterAtPos3 THEN #StateNo := 320; END_IF;
END_REGION

REGION Network 86: Actions for STATE Num:320 StWtLifterAtPos3
   RUNG wire#powerrail
      Contact( #sStWtLifterAtPos3 )
      Coil( #qLifterAtPos3 )
   END_RUNG
   // the same network as SCL:
   #qLifterAtPos3 := #sStWtLifterAtPos3;
END_REGION

REGION Network 87: Transition for STATE Num:330 StWtL2S1Down
   RUNG wire#powerrail
      Contact( #sStWtL2S1Down )
      I_Contact( #sStWtResetRel )
      Contact( #sSst )
      Contact( #iL2S1Down )
      Coil( #sStWtL2S1Down_T1 )
   END_RUNG
   // the same network as SCL:
   #sStWtL2S1Down_T1 := #sStWtL2S1Down AND NOT #sStWtResetRel AND #sSst AND #iL2S1Down;
END_REGION

REGION Network 88: STATE Num:330 StWtL2S1Down
   RUNG wire#powerrail
      Contact( #sStWtL2S1Down )
      wire#w1
      I_Contact( #sStWtResetRel )
      I_Contact( #sStWtL2S1Down_T1 )
      wire#w2
      Coil( #sStWtL2S1Down )
   END_RUNG
   RUNG wire#powerrail
      Contact( #sStWtLifterAtPos3_T1 )
   END_RUNG wire#w1
   RUNG wire#powerrail
      Contact( #sStRecovery_T6 )
   END_RUNG wire#w1
   RUNG wire#w2
      { S7_GenerateENO := "TRUE" } Move(in := 330, out1 => #StateNo)
   END_RUNG
   // the same network as SCL:
   #sStWtL2S1Down := (#sStWtL2S1Down OR #sStWtLifterAtPos3_T1 OR #sStRecovery_T6) AND NOT #sStWtResetRel AND NOT #sStWtL2S1Down_T1;
   IF #sStWtL2S1Down THEN #StateNo := 330; END_IF;
END_REGION

REGION Network 89: Actions for STATE Num:330 StWtL2S1Down
   RUNG wire#powerrail
      Contact( #sStWtL2S1Down )
      Coil( #qL1S1Down )
   END_RUNG
   // the same network as SCL:
   #qL1S1Down := #sStWtL2S1Down;
END_REGION

REGION Network 90: Transition for STATE Num:340 StWtOTSFrmTT
   RUNG wire#powerrail
      Contact( #sStWtOTSFrmTT )
      I_Contact( #sStWtResetRel )
      Contact( #sSst )
      Contact( #iOTSFrmConv )
      Coil( #sStWtOTSFrmTT_T1 )
   END_RUNG
   // the same network as SCL:
   #sStWtOTSFrmTT_T1 := #sStWtOTSFrmTT AND NOT #sStWtResetRel AND #sSst AND #iOTSFrmConv;
END_REGION

REGION Network 91: STATE Num:340 StWtOTSFrmTT
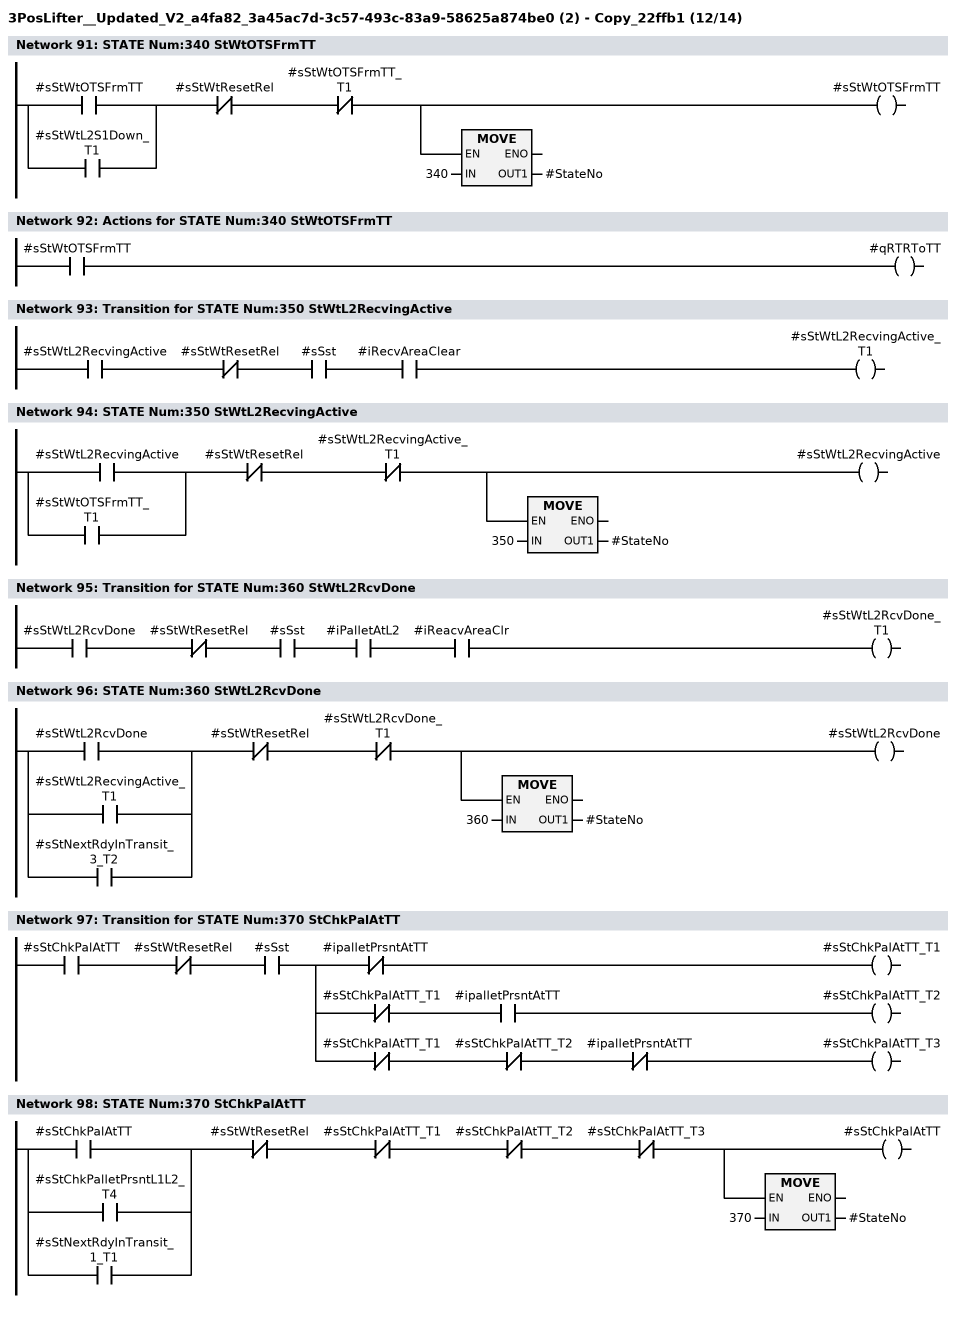
   RUNG wire#powerrail
      Contact( #sStWtOTSFrmTT )
      wire#w1
      I_Contact( #sStWtResetRel )
      I_Contact( #sStWtOTSFrmTT_T1 )
      wire#w2
      Coil( #sStWtOTSFrmTT )
   END_RUNG
   RUNG wire#powerrail
      Contact( #sStWtL2S1Down_T1 )
   END_RUNG wire#w1
   RUNG wire#w2
      { S7_GenerateENO := "TRUE" } Move(in := 340, out1 => #StateNo)
   END_RUNG
   // the same network as SCL:
   #sStWtOTSFrmTT := (#sStWtOTSFrmTT OR #sStWtL2S1Down_T1) AND NOT #sStWtResetRel AND NOT #sStWtOTSFrmTT_T1;
   IF #sStWtOTSFrmTT THEN #StateNo := 340; END_IF;
END_REGION

REGION Network 92: Actions for STATE Num:340 StWtOTSFrmTT
   RUNG wire#powerrail
      Contact( #sStWtOTSFrmTT )
      Coil( #qRTRToTT )
   END_RUNG
   // the same network as SCL:
   #qRTRToTT := #sStWtOTSFrmTT;
END_REGION

REGION Network 93: Transition for STATE Num:350 StWtL2RecvingActive
   RUNG wire#powerrail
      Contact( #sStWtL2RecvingActive )
      I_Contact( #sStWtResetRel )
      Contact( #sSst )
      Contact( #iRecvAreaClear )
      Coil( #sStWtL2RecvingActive_T1 )
   END_RUNG
   // the same network as SCL:
   #sStWtL2RecvingActive_T1 := #sStWtL2RecvingActive AND NOT #sStWtResetRel AND #sSst AND #iRecvAreaClear;
END_REGION

REGION Network 94: STATE Num:350 StWtL2RecvingActive
   RUNG wire#powerrail
      Contact( #sStWtL2RecvingActive )
      wire#w1
      I_Contact( #sStWtResetRel )
      I_Contact( #sStWtL2RecvingActive_T1 )
      wire#w2
      Coil( #sStWtL2RecvingActive )
   END_RUNG
   RUNG wire#powerrail
      Contact( #sStWtOTSFrmTT_T1 )
   END_RUNG wire#w1
   RUNG wire#w2
      { S7_GenerateENO := "TRUE" } Move(in := 350, out1 => #StateNo)
   END_RUNG
   // the same network as SCL:
   #sStWtL2RecvingActive := (#sStWtL2RecvingActive OR #sStWtOTSFrmTT_T1) AND NOT #sStWtResetRel AND NOT #sStWtL2RecvingActive_T1;
   IF #sStWtL2RecvingActive THEN #StateNo := 350; END_IF;
END_REGION

REGION Network 95: Transition for STATE Num:360 StWtL2RcvDone
   RUNG wire#powerrail
      Contact( #sStWtL2RcvDone )
      I_Contact( #sStWtResetRel )
      Contact( #sSst )
      Contact( #iPalletAtL2 )
      Contact( #iReacvAreaClr )
      Coil( #sStWtL2RcvDone_T1 )
   END_RUNG
   // the same network as SCL:
   #sStWtL2RcvDone_T1 := #sStWtL2RcvDone AND NOT #sStWtResetRel AND #sSst AND #iPalletAtL2 AND #iReacvAreaClr;
END_REGION

REGION Network 96: STATE Num:360 StWtL2RcvDone
   RUNG wire#powerrail
      Contact( #sStWtL2RcvDone )
      wire#w1
      I_Contact( #sStWtResetRel )
      I_Contact( #sStWtL2RcvDone_T1 )
      wire#w2
      Coil( #sStWtL2RcvDone )
   END_RUNG
   RUNG wire#powerrail
      Contact( #sStWtL2RecvingActive_T1 )
   END_RUNG wire#w1
   RUNG wire#powerrail
      Contact( #sStNextRdyInTransit_3_T2 )
   END_RUNG wire#w1
   RUNG wire#w2
      { S7_GenerateENO := "TRUE" } Move(in := 360, out1 => #StateNo)
   END_RUNG
   // the same network as SCL:
   #sStWtL2RcvDone := (#sStWtL2RcvDone OR #sStWtL2RecvingActive_T1 OR #sStNextRdyInTransit_3_T2) AND NOT #sStWtResetRel AND NOT #sStWtL2RcvDone_T1;
   IF #sStWtL2RcvDone THEN #StateNo := 360; END_IF;
END_REGION

REGION Network 97: Transition for STATE Num:370 StChkPalAtTT
   RUNG wire#powerrail
      Contact( #sStChkPalAtTT )
      I_Contact( #sStWtResetRel )
      Contact( #sSst )
      wire#w1
      I_Contact( #ipalletPrsntAtTT )
      Coil( #sStChkPalAtTT_T1 )
   END_RUNG
   RUNG wire#w1
      I_Contact( #sStChkPalAtTT_T1 )
      Contact( #ipalletPrsntAtTT )
      Coil( #sStChkPalAtTT_T2 )
   END_RUNG
   RUNG wire#w1
      I_Contact( #sStChkPalAtTT_T1 )
      I_Contact( #sStChkPalAtTT_T2 )
      I_Contact( #ipalletPrsntAtTT )
      Coil( #sStChkPalAtTT_T3 )
   END_RUNG
   // the same network as SCL:
   #_w1 := #sStChkPalAtTT AND NOT #sStWtResetRel AND #sSst;
   #sStChkPalAtTT_T1 := #_w1 AND NOT #ipalletPrsntAtTT;
   #sStChkPalAtTT_T2 := #_w1 AND NOT #sStChkPalAtTT_T1 AND #ipalletPrsntAtTT;
   #sStChkPalAtTT_T3 := #_w1 AND NOT #sStChkPalAtTT_T1 AND NOT #sStChkPalAtTT_T2 AND NOT #ipalletPrsntAtTT;
END_REGION

REGION Network 98: STATE Num:370 StChkPalAtTT
   RUNG wire#powerrail
      Contact( #sStChkPalAtTT )
      wire#w1
      I_Contact( #sStWtResetRel )
      I_Contact( #sStChkPalAtTT_T1 )
      I_Contact( #sStChkPalAtTT_T2 )
      I_Contact( #sStChkPalAtTT_T3 )
      wire#w2
      Coil( #sStChkPalAtTT )
   END_RUNG
   RUNG wire#powerrail
      Contact( #sStChkPalletPrsntL1L2_T4 )
   END_RUNG wire#w1
   RUNG wire#powerrail
      Contact( #sStNextRdyInTransit_1_T1 )
   END_RUNG wire#w1
   RUNG wire#w2
      { S7_GenerateENO := "TRUE" } Move(in := 370, out1 => #StateNo)
   END_RUNG
   // the same network as SCL:
   #sStChkPalAtTT := (#sStChkPalAtTT OR #sStChkPalletPrsntL1L2_T4 OR #sStNextRdyInTransit_1_T1) AND NOT #sStWtResetRel AND NOT #sStChkPalAtTT_T1 AND NOT #sStChkPalAtTT_T2 AND NOT #sStChkPalAtTT_T3;
   IF #sStChkPalAtTT THEN #StateNo := 370; END_IF;
END_REGION

REGION Network 99: Transition for STATE Num:380 StWtLifterAtPos2
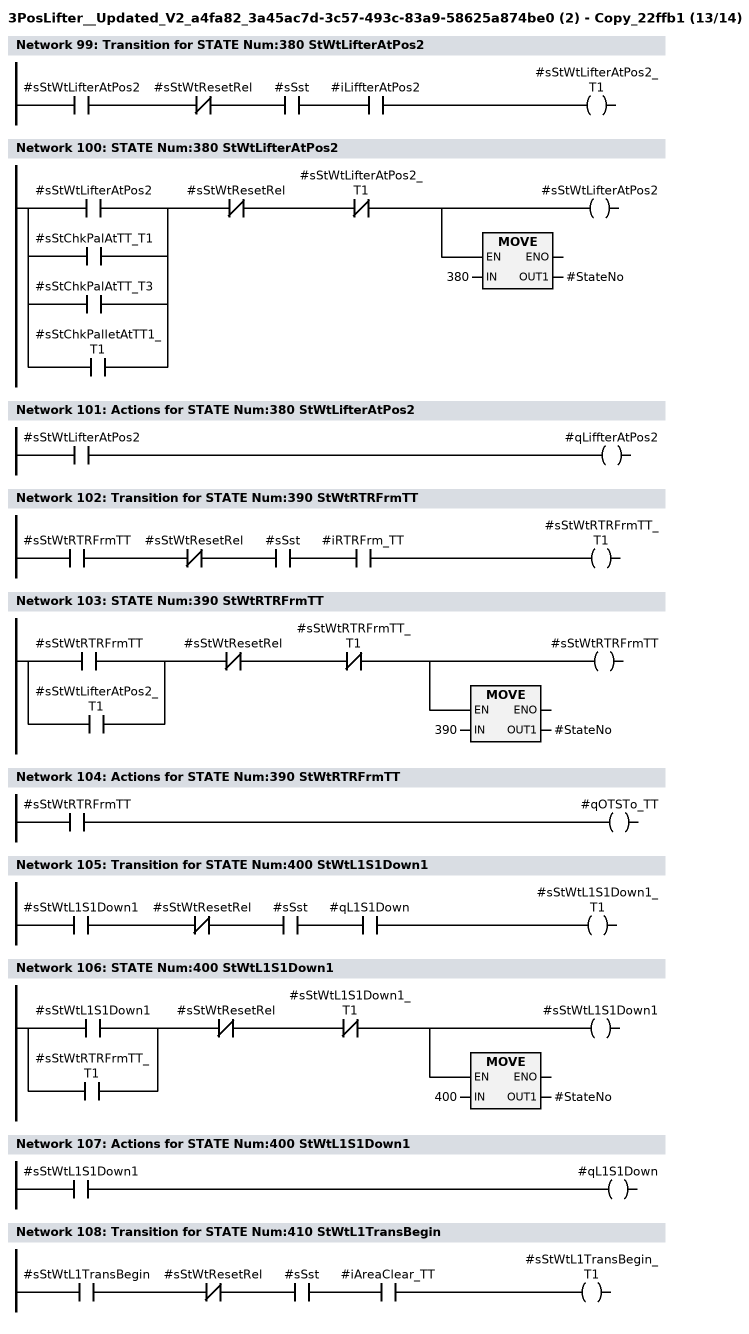
   RUNG wire#powerrail
      Contact( #sStWtLifterAtPos2 )
      I_Contact( #sStWtResetRel )
      Contact( #sSst )
      Contact( #iLiffterAtPos2 )
      Coil( #sStWtLifterAtPos2_T1 )
   END_RUNG
   // the same network as SCL:
   #sStWtLifterAtPos2_T1 := #sStWtLifterAtPos2 AND NOT #sStWtResetRel AND #sSst AND #iLiffterAtPos2;
END_REGION

REGION Network 100: STATE Num:380 StWtLifterAtPos2
   RUNG wire#powerrail
      Contact( #sStWtLifterAtPos2 )
      wire#w1
      I_Contact( #sStWtResetRel )
      I_Contact( #sStWtLifterAtPos2_T1 )
      wire#w2
      Coil( #sStWtLifterAtPos2 )
   END_RUNG
   RUNG wire#powerrail
      Contact( #sStChkPalAtTT_T1 )
   END_RUNG wire#w1
   RUNG wire#powerrail
      Contact( #sStChkPalAtTT_T3 )
   END_RUNG wire#w1
   RUNG wire#powerrail
      Contact( #sStChkPalletAtTT1_T1 )
   END_RUNG wire#w1
   RUNG wire#w2
      { S7_GenerateENO := "TRUE" } Move(in := 380, out1 => #StateNo)
   END_RUNG
   // the same network as SCL:
   #sStWtLifterAtPos2 := (#sStWtLifterAtPos2 OR #sStChkPalAtTT_T1 OR #sStChkPalAtTT_T3 OR #sStChkPalletAtTT1_T1) AND NOT #sStWtResetRel AND NOT #sStWtLifterAtPos2_T1;
   IF #sStWtLifterAtPos2 THEN #StateNo := 380; END_IF;
END_REGION

REGION Network 101: Actions for STATE Num:380 StWtLifterAtPos2
   RUNG wire#powerrail
      Contact( #sStWtLifterAtPos2 )
      Coil( #qLiffterAtPos2 )
   END_RUNG
   // the same network as SCL:
   #qLiffterAtPos2 := #sStWtLifterAtPos2;
END_REGION

REGION Network 102: Transition for STATE Num:390 StWtRTRFrmTT
   RUNG wire#powerrail
      Contact( #sStWtRTRFrmTT )
      I_Contact( #sStWtResetRel )
      Contact( #sSst )
      Contact( #iRTRFrm_TT )
      Coil( #sStWtRTRFrmTT_T1 )
   END_RUNG
   // the same network as SCL:
   #sStWtRTRFrmTT_T1 := #sStWtRTRFrmTT AND NOT #sStWtResetRel AND #sSst AND #iRTRFrm_TT;
END_REGION

REGION Network 103: STATE Num:390 StWtRTRFrmTT
   RUNG wire#powerrail
      Contact( #sStWtRTRFrmTT )
      wire#w1
      I_Contact( #sStWtResetRel )
      I_Contact( #sStWtRTRFrmTT_T1 )
      wire#w2
      Coil( #sStWtRTRFrmTT )
   END_RUNG
   RUNG wire#powerrail
      Contact( #sStWtLifterAtPos2_T1 )
   END_RUNG wire#w1
   RUNG wire#w2
      { S7_GenerateENO := "TRUE" } Move(in := 390, out1 => #StateNo)
   END_RUNG
   // the same network as SCL:
   #sStWtRTRFrmTT := (#sStWtRTRFrmTT OR #sStWtLifterAtPos2_T1) AND NOT #sStWtResetRel AND NOT #sStWtRTRFrmTT_T1;
   IF #sStWtRTRFrmTT THEN #StateNo := 390; END_IF;
END_REGION

REGION Network 104: Actions for STATE Num:390 StWtRTRFrmTT
   RUNG wire#powerrail
      Contact( #sStWtRTRFrmTT )
      Coil( #qOTSTo_TT )
   END_RUNG
   // the same network as SCL:
   #qOTSTo_TT := #sStWtRTRFrmTT;
END_REGION

REGION Network 105: Transition for STATE Num:400 StWtL1S1Down1
   RUNG wire#powerrail
      Contact( #sStWtL1S1Down1 )
      I_Contact( #sStWtResetRel )
      Contact( #sSst )
      Contact( #qL1S1Down )
      Coil( #sStWtL1S1Down1_T1 )
   END_RUNG
   // the same network as SCL:
   #sStWtL1S1Down1_T1 := #sStWtL1S1Down1 AND NOT #sStWtResetRel AND #sSst AND #qL1S1Down;
END_REGION

REGION Network 106: STATE Num:400 StWtL1S1Down1
   RUNG wire#powerrail
      Contact( #sStWtL1S1Down1 )
      wire#w1
      I_Contact( #sStWtResetRel )
      I_Contact( #sStWtL1S1Down1_T1 )
      wire#w2
      Coil( #sStWtL1S1Down1 )
   END_RUNG
   RUNG wire#powerrail
      Contact( #sStWtRTRFrmTT_T1 )
   END_RUNG wire#w1
   RUNG wire#w2
      { S7_GenerateENO := "TRUE" } Move(in := 400, out1 => #StateNo)
   END_RUNG
   // the same network as SCL:
   #sStWtL1S1Down1 := (#sStWtL1S1Down1 OR #sStWtRTRFrmTT_T1) AND NOT #sStWtResetRel AND NOT #sStWtL1S1Down1_T1;
   IF #sStWtL1S1Down1 THEN #StateNo := 400; END_IF;
END_REGION

REGION Network 107: Actions for STATE Num:400 StWtL1S1Down1
   RUNG wire#powerrail
      Contact( #sStWtL1S1Down1 )
      Coil( #qL1S1Down )
   END_RUNG
   // the same network as SCL:
   #qL1S1Down := #sStWtL1S1Down1;
END_REGION

REGION Network 108: Transition for STATE Num:410 StWtL1TransBegin
   RUNG wire#powerrail
      Contact( #sStWtL1TransBegin )
      I_Contact( #sStWtResetRel )
      Contact( #sSst )
      Contact( #iAreaClear_TT )
      Coil( #sStWtL1TransBegin_T1 )
   END_RUNG
   // the same network as SCL:
   #sStWtL1TransBegin_T1 := #sStWtL1TransBegin AND NOT #sStWtResetRel AND #sSst AND #iAreaClear_TT;
END_REGION

REGION Network 109: STATE Num:410 StWtL1TransBegin
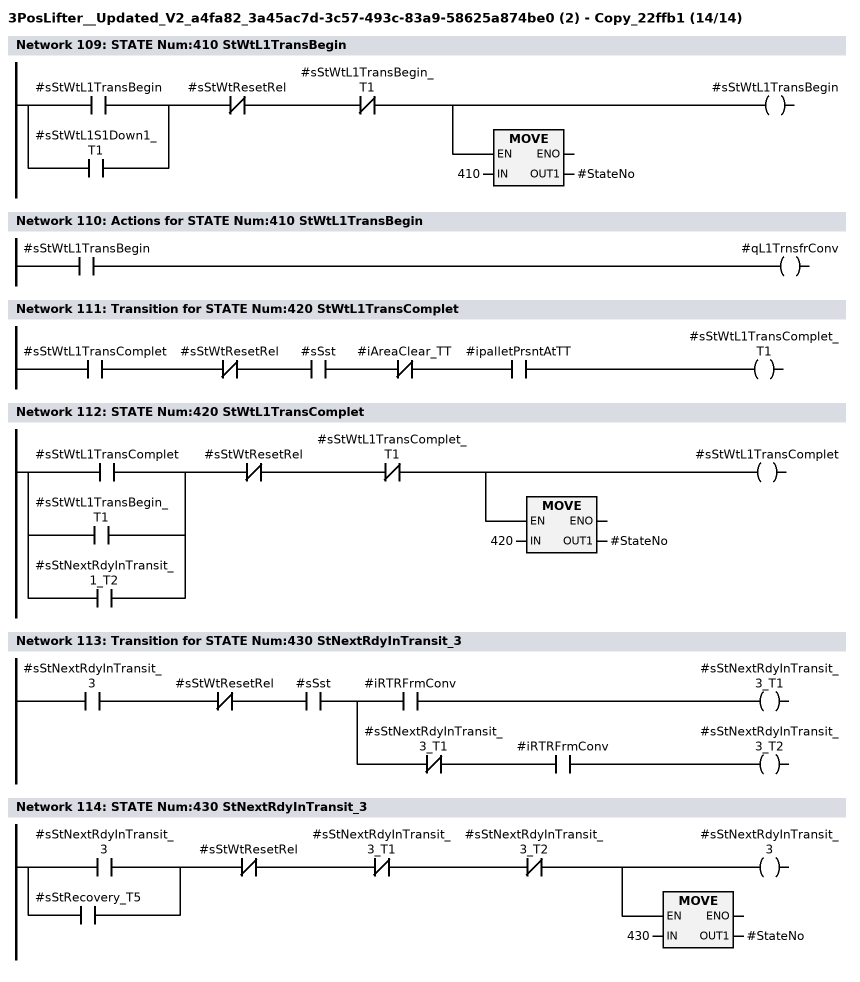
   RUNG wire#powerrail
      Contact( #sStWtL1TransBegin )
      wire#w1
      I_Contact( #sStWtResetRel )
      I_Contact( #sStWtL1TransBegin_T1 )
      wire#w2
      Coil( #sStWtL1TransBegin )
   END_RUNG
   RUNG wire#powerrail
      Contact( #sStWtL1S1Down1_T1 )
   END_RUNG wire#w1
   RUNG wire#w2
      { S7_GenerateENO := "TRUE" } Move(in := 410, out1 => #StateNo)
   END_RUNG
   // the same network as SCL:
   #sStWtL1TransBegin := (#sStWtL1TransBegin OR #sStWtL1S1Down1_T1) AND NOT #sStWtResetRel AND NOT #sStWtL1TransBegin_T1;
   IF #sStWtL1TransBegin THEN #StateNo := 410; END_IF;
END_REGION

REGION Network 110: Actions for STATE Num:410 StWtL1TransBegin
   RUNG wire#powerrail
      Contact( #sStWtL1TransBegin )
      Coil( #qL1TrnsfrConv )
   END_RUNG
   // the same network as SCL:
   #qL1TrnsfrConv := #sStWtL1TransBegin;
END_REGION

REGION Network 111: Transition for STATE Num:420 StWtL1TransComplet
   RUNG wire#powerrail
      Contact( #sStWtL1TransComplet )
      I_Contact( #sStWtResetRel )
      Contact( #sSst )
      I_Contact( #iAreaClear_TT )
      Contact( #ipalletPrsntAtTT )
      Coil( #sStWtL1TransComplet_T1 )
   END_RUNG
   // the same network as SCL:
   #sStWtL1TransComplet_T1 := #sStWtL1TransComplet AND NOT #sStWtResetRel AND #sSst AND NOT #iAreaClear_TT AND #ipalletPrsntAtTT;
END_REGION

REGION Network 112: STATE Num:420 StWtL1TransComplet
   RUNG wire#powerrail
      Contact( #sStWtL1TransComplet )
      wire#w1
      I_Contact( #sStWtResetRel )
      I_Contact( #sStWtL1TransComplet_T1 )
      wire#w2
      Coil( #sStWtL1TransComplet )
   END_RUNG
   RUNG wire#powerrail
      Contact( #sStWtL1TransBegin_T1 )
   END_RUNG wire#w1
   RUNG wire#powerrail
      Contact( #sStNextRdyInTransit_1_T2 )
   END_RUNG wire#w1
   RUNG wire#w2
      { S7_GenerateENO := "TRUE" } Move(in := 420, out1 => #StateNo)
   END_RUNG
   // the same network as SCL:
   #sStWtL1TransComplet := (#sStWtL1TransComplet OR #sStWtL1TransBegin_T1 OR #sStNextRdyInTransit_1_T2) AND NOT #sStWtResetRel AND NOT #sStWtL1TransComplet_T1;
   IF #sStWtL1TransComplet THEN #StateNo := 420; END_IF;
END_REGION

REGION Network 113: Transition for STATE Num:430 StNextRdyInTransit_3
   RUNG wire#powerrail
      Contact( #sStNextRdyInTransit_3 )
      I_Contact( #sStWtResetRel )
      Contact( #sSst )
      wire#w1
      Contact( #iRTRFrmConv )
      Coil( #sStNextRdyInTransit_3_T1 )
   END_RUNG
   RUNG wire#w1
      I_Contact( #sStNextRdyInTransit_3_T1 )
      Contact( #iRTRFrmConv )
      Coil( #sStNextRdyInTransit_3_T2 )
   END_RUNG
   // the same network as SCL:
   #_w1 := #sStNextRdyInTransit_3 AND NOT #sStWtResetRel AND #sSst;
   #sStNextRdyInTransit_3_T1 := #_w1 AND #iRTRFrmConv;
   #sStNextRdyInTransit_3_T2 := #_w1 AND NOT #sStNextRdyInTransit_3_T1 AND #iRTRFrmConv;
END_REGION

REGION Network 114: STATE Num:430 StNextRdyInTransit_3
   RUNG wire#powerrail
      Contact( #sStNextRdyInTransit_3 )
      wire#w1
      I_Contact( #sStWtResetRel )
      I_Contact( #sStNextRdyInTransit_3_T1 )
      I_Contact( #sStNextRdyInTransit_3_T2 )
      wire#w2
      Coil( #sStNextRdyInTransit_3 )
   END_RUNG
   RUNG wire#powerrail
      Contact( #sStRecovery_T5 )
   END_RUNG wire#w1
   RUNG wire#w2
      { S7_GenerateENO := "TRUE" } Move(in := 430, out1 => #StateNo)
   END_RUNG
   // the same network as SCL:
   #sStNextRdyInTransit_3 := (#sStNextRdyInTransit_3 OR #sStRecovery_T5) AND NOT #sStWtResetRel AND NOT #sStNextRdyInTransit_3_T1 AND NOT #sStNextRdyInTransit_3_T2;
   IF #sStNextRdyInTransit_3 THEN #StateNo := 430; END_IF;
END_REGION
END_FUNCTION_BLOCK
